// TwinCAT 3 PLC project TC3_Tester_Palet
// ProgramVersion: 3.1.4026.26
// libraries:
//   Tc2_Standard, * (Beckhoff Automation GmbH)
//   Tc2_System, * (Beckhoff Automation GmbH)
// project tree:
//   DUTs/DUTs/ E_StackAlarm.TcDUT, ST_StackCfg.TcDUT, ST_StackMem.TcDUT, ST_StackPersist.TcDUT, ST_St04Cfg.TcDUT, ST_St04_In.TcDUT, ST_St04_Out.TcDUT, ST_St05Cfg.TcDUT, ST_St05_In.TcDUT, ST_St05_Out.TcDUT, E_CylAlarm.TcDUT, E_CylFeedback.TcDUT, E_CylState.TcDUT, E_CylValve.TcDUT, ST_CylCfg.TcDUT, ST_CylMem.TcDUT, ST_CylPersist.TcDUT, E_MachineMode.TcDUT, E_NodeAlarm.TcDUT, E_NodeState.TcDUT, E_WaitCause.TcDUT, ST_ConvCfg.TcDUT, ST_ConvMem.TcDUT, ST_ConvPersist.TcDUT, E_NordSK550P_State.TcDUT, ST_NordSK550P_In.TcDUT, ST_NordSK550P_Out.TcDUT
//   POUs/POUs/FB/ FB_StackLift.TcPOU, FB_Station03_Destack.TcPOU, FB_Station11_Stack.TcPOU, FB_Station04_Press.TcPOU, FB_Station05_Tear.TcPOU, FB_CylPosMonitor.TcPOU, FB_CamAxis.TcPOU, FB_CsvLogger.TcPOU, FB_Cylinder.TcPOU, FB_RollerConveyor.TcPOU, FB_TransportNodeBase.TcPOU, FB_StationPickup.TcPOU, FB_NordSK550PP.TcPOU, TestFb.TcPOU
//   GVLs/ GVL_PERSIST.TcGVL, GVL.TcGVL, GVL_IO.TcGVL, GVL_SAFETY.TcGVL
//   / PlcTask.TcTTO
//   POUs/ PRG_Machine.TcPOU, MAIN.TcPOU

CONFIGURATION TC3_Tester_Palet
    RESOURCE PLC ON TwinCAT3
        TASK PlcTask(INTERVAL := T#10ms, PRIORITY := 20);
        PROGRAM MAIN WITH PlcTask : MAIN;
    END_RESOURCE
END_CONFIGURATION

// ---- DUTs/DUTs/E_StackAlarm.TcDUT
TYPE E_StackAlarm :
(
	ALM_STK_NONE			:= 0,

	// Wozek nie dojechal do pozycji w zadanym czasie
	ALM_STK_MOVE_TIMEOUT	:= 1,

	// Szczeki nie potwierdzily ruchu
	ALM_STK_JAW_TIMEOUT		:= 2,

	// Pozycje wpisane przez operatora nie tworza rosnacego
	// ani malejacego ciagu - dol / srodek / gora musza lezec
	// po kolei, inaczej wozek pojechalby w zla strone
	ALM_STK_POS_INVALID		:= 3,

	// Blad falownika wozka
	ALM_STK_DRIVE_FAULT		:= 4,

	// Brak wywolania M_Config
	ALM_STK_NOT_CONFIGURED	:= 5,

	// Wozek zjechal z potwierdzonej pozycji bez komendy
	ALM_STK_POSITION_LOST	:= 6
);
END_TYPE

// ---- DUTs/DUTs/ST_StackCfg.TcDUT
TYPE ST_StackCfg :
STRUCT
	// =========================================================
	// DESZTAPLARKA / SZTAPLARKA - NASTAWY NIEULOTNE
	// =========================================================
	//
	// Obie maszyny maja te sama kinematyke: wozek ze szczekami
	// jezdzacy w pionie na falowniku, z enkoderem absolutnym,
	// i trzy pozycje robocze. Rozni je tylko kolejnosc krokow.
	//
	// ---------------------------------------------------------
	// TRZY POZYCJE
	// ---------------------------------------------------------
	// Liczac od dolu, przy stosie stojacym na transporterze:
	//
	//   diPosBottom  wysokosc desek PIERWSZEJ palety od dolu
	//   diPosMiddle  wysokosc desek DRUGIEJ palety od dolu
	//   diPosTop     pozycja stosu uniesionego
	//
	// Desztaplarka chwyta na diPosMiddle - czyli pod druga
	// palete - i jedzie na diPosTop, przez co najnizsza paleta
	// zostaje na transporterze. Odklada stos na diPosBottom.
	//
	// Sztaplarka odklada trzymany stos na diPosMiddle, czyli
	// wprost na palete, ktora wlasnie przyjechala, a chwyta
	// caly stos od spodu na diPosBottom.
	//
	// Wartosci wpisuje operator z palca. Automat bazujacy
	// dopiszemy pozniej - dlatego jest kontrola poprawnosci:
	// trzy pozycje musza tworzyc ciag rosnacy albo malejacy.

	sName				: STRING(31);

	// Wartosci dobrane na maszynie. Enkoder jednoobrotowy
	// 0..65535, zero na pozycji DOLNEJ. Obie maszyny maja na
	// razie te same punkty.
	//
	// UWAGA: to sa wartosci NIEULOTNE. Wpis z deklaracji
	// obowiazuje tylko przy pierwszym pobraniu projektu albo
	// po skasowaniu danych nieulotnych. Pozniejsza zmiana tej
	// liczby w kodzie nie ruszy nastawy na sterowniku - trzeba
	// ja poprawic online albo zrobic "Reset origin".
	diPosBottom			: DINT := 0;
	diPosMiddle			: DINT := 16000;
	diPosTop			: DINT := 24000;

	// Okno, w ktorym uznajemy pozycje za osiagnieta
	diWindow			: DINT := 20;

	// Odleglosc, od ktorej zwalniamy do predkosci dojazdowej
	diSlowZone			: DINT := 300;

	// TRUE = rosnaca wartosc enkodera odpowiada jezdzie
	// napedem DO PRZODU
	xIncreaseIsForward	: BOOL := TRUE;


	// ---------------------------------------------------------
	// PREDKOSCI I CZASY
	// ---------------------------------------------------------

	lrFreqFast			: LREAL := 35.0;
	lrFreqSlow			: LREAL := 10.0;
	lrFreqManual		: LREAL := 8.0;

	// Czas, w ktorym wozek musi dojechac do pozycji
	tMoveWatchdog		: TIME := T#15S;

	// Uspokojenie po dojezdzie, zanim ruszymy szczekami
	tSettle				: TIME := T#200MS;


	// ---------------------------------------------------------
	// STOS
	// ---------------------------------------------------------
	//
	// Na razie stala liczba palet w stosie. Czujnik wykrywajacy,
	// ze wszystkie palety zostaly wydane, dojdzie pozniej -
	// wtedy ta wartosc bedzie tylko wartoscia oczekiwana.

	nStackSize			: INT := 15;

END_STRUCT
END_TYPE

// ---- DUTs/DUTs/ST_StackMem.TcDUT
TYPE ST_StackMem :
STRUCT
	// =========================================================
	// PAMIEC DESZTAPLARKI / SZTAPLARKI - ZMIENNE NIEULOTNE
	// =========================================================
	//
	// Po zaniku zasilania maszyna musi wiedziec, ile palet
	// zostalo w stosie i ile wisi na szczekach. Bez tego
	// operator musialby rozladowac stacje recznie.

	// Stos dojechal na stacje i zostal potwierdzony czujnikami
	xStackArrived	: BOOL;

	// DESZTAPLARKA: ile palet zostalo do wydania, wliczajac te,
	// ktora aktualnie lezy na transporterze
	nRemaining		: INT;

	// SZTAPLARKA: ile palet wisi na szczekach
	nHeld			: INT;

	// Szczeki trzymaja ladunek - po zaniku zasilania nie wolno
	// ich otworzyc bez sprowadzenia wozka na pozycje odkladania
	xJawsLoaded		: BOOL;

	// Ostatnia znana pozycja enkodera, zapisywana na biezaco.
	// Po starcie porownujemy ja z odczytem: jesli sie zgadza,
	// enkoder utrzymal wartosc przez zanik zasilania i NIE ma
	// potrzeby bazowania. Jesli nie - kod sam to zglosi.
	diLastPos		: DINT;

	// TRUE = po starcie odczyt enkodera nie zgodzil sie
	// z zapamietanym. Trzeba zbazowac pozycje dolna.
	xNeedHoming		: BOOL;

END_STRUCT
END_TYPE

// ---- DUTs/DUTs/ST_StackPersist.TcDUT
TYPE ST_StackPersist :
STRUCT
	Cfg		: ST_StackCfg;
	Mem		: ST_StackMem;
END_STRUCT
END_TYPE

// ---- DUTs/DUTs/ST_St04Cfg.TcDUT
TYPE ST_St04Cfg :
STRUCT
	// =========================================================
	// STACJA 4 - TEST SCISKANIA, NASTAWY NIEULOTNE
	// =========================================================
	//
	// Test toczy sie na JADACEJ palecie. Rolki dociskowe kreca
	// sie caly czas, a silowniki napieraja na deski w trakcie
	// przejazdu. Dlatego przerwanie uniewaznia wynik -
	// aConv[4].Cfg.xNokOnInterrupt musi byc TRUE.

	// ---------------------------------------------------------
	// CZUJNIK WSTEPNY
	// ---------------------------------------------------------
	//
	// Czujnik przed stacja, od ktorego liczy sie czas do wysuwu
	// silownikow. Na dzien pisania kodu jeszcze nie zamontowany.
	//
	// xPreSensorInstalled = FALSE: czasowka startuje od chwili
	// ruszenia palety z poprzedniej stacji (tEntryToUpper).
	// Po montazu wystarczy przelaczyc bit - kod sie nie zmienia.

	xPreSensorInstalled	: BOOL := FALSE;

	// TRUE = logika odwrocona, tak jak czujniki koncowe
	// (0 na wejsciu = czujnik cos widzi)
	xPreSensorInverted	: BOOL := TRUE;


	// ---------------------------------------------------------
	// CZASY SEKWENCJI
	// ---------------------------------------------------------

	// Od czujnika wstepnego do wysuwu silownikow GORNYCH
	tPreToUpper			: TIME := T#500MS;

	// To samo, gdy czujnika wstepnego jeszcze nie ma -
	// liczone od rozpoczecia wjazdu
	tEntryToUpper		: TIME := T#3S;

	// Od wysuwu gornych do wysuwu DOLNYCH.
	// Gorne ida pierwsze, zeby dolne nie uniosly palety,
	// ale odstep ma byc symboliczny - dociski maja isc razem.
	tUpperToLower		: TIME := T#100MS;

	// Watchdog calej operacji
	tOpWatchdog			: TIME := T#60S;


	// ---------------------------------------------------------
	// ROLKI DOCISKOWE
	// ---------------------------------------------------------
	//
	// Falownik 3. Rolki na koncach silownikow gornych sa
	// napedzane, zeby paleta nie utknela pod dociskiem.

	lrRollerFreq		: LREAL := 25.0;

END_STRUCT
END_TYPE

// ---- DUTs/DUTs/ST_St04_In.TcDUT
TYPE ST_St04_In :
STRUCT
	// =========================================================
	// STACJA 4 - SYGNALY WEJSCIOWE
	// =========================================================

	// Czujnik wstepny - jeszcze niepodlinkowany.
	// Do czasu montazu zostawic Cfg.xPreSensorInstalled = FALSE.
	xPreSensRaw		: BOOL := TRUE;

	// Przetworniki polozenia IO-Link, po jednym na KAZDY
	// silownik, mimo ze zawory steruja grupami:
	//   1..3  dolne
	//   4..6  gorne od szerokich desek
	//   7..8  gorne od waskich desek
	adiCylPos		: ARRAY[1..8] OF DINT;

END_STRUCT
END_TYPE

// ---- DUTs/DUTs/ST_St04_Out.TcDUT
TYPE ST_St04_Out :
STRUCT
	// =========================================================
	// STACJA 4 - CEWKI ZAWOROW
	// =========================================================
	//
	// Mapowanie w MAIN wg opisu wyjsc:
	//   xLowerExtend        -> GVL.OUTPUTS[4]   dolne wysun
	//   xLowerRetract       -> GVL.OUTPUTS[3]   dolne cofnij
	//   xUpperWideExtend    -> GVL.OUTPUTS[7]   gorne zewnetrzne
	//                                           i srodkowa wysun
	//   xUpperWideRetract   -> GVL.OUTPUTS[2]   te same cofnij
	//   xUpperNarrowExtend  -> GVL.OUTPUTS[5]   gorne srodkowe wysun
	//   xUpperNarrowRetract -> GVL.OUTPUTS[6]   gorne srodkowe cofnij
	//
	// [?] Opis wyjsc 2/7 i 5/6 nazywa obie grupy "srodkowymi".
	// Przyjete: 7/2 to trzy silowniki od szerokich desek,
	// 5/6 to dwa od waskich. Do potwierdzenia na maszynie -
	// zamiana dotyczy wylacznie mapowania w MAIN, nie kodu stacji.

	xLowerExtend		: BOOL;
	xLowerRetract		: BOOL;

	xUpperWideExtend	: BOOL;
	xUpperWideRetract	: BOOL;

	xUpperNarrowExtend	: BOOL;
	xUpperNarrowRetract	: BOOL;

END_STRUCT
END_TYPE

// ---- DUTs/DUTs/ST_St05Cfg.TcDUT
TYPE ST_St05Cfg :
STRUCT
	// =========================================================
	// STACJA 5 - TEST ROZRYWANIA, NASTAWY NIEULOTNE
	// =========================================================
	//
	// Czasy samych ruchow silownikow siedza w ich wlasnych
	// rekordach (GVL_PERSIST.aCyl). Tutaj sa tylko czasy
	// nalezace do SEKWENCJI stacji.

	// Od potwierdzenia palety na blokadzie do podniesienia szczek
	tDetectToLift		: TIME := T#500MS;

	// Od zamkniecia szczek do rozpoczecia rozrywania
	tJawsToPull			: TIME := T#300MS;

	// Watchdog calej operacji testu
	tOpWatchdog			: TIME := T#60S;

	// UWAGA: blokada NIE podnosi sie na czasowke. Idzie w gore
	// w chwili, gdy z poprzedniej stacji rusza paleta - wtedy
	// nikt jej nie stoi na drodze, a czasu na podniesienie jest
	// tyle, ile trwa przejazd. Czas ruchu samej blokady i jego
	// watchdog siedza w GVL_PERSIST.aCyl.

END_STRUCT
END_TYPE

// ---- DUTs/DUTs/ST_St05_In.TcDUT
TYPE ST_St05_In :
STRUCT
	// =========================================================
	// STACJA 5 - SYGNALY WEJSCIOWE
	// =========================================================
	//
	// Cale mapowanie z GVL siedzi w jednym miejscu w MAIN.
	// Blok stacji nie siega do GVL bezposrednio.

	// Blokada punktu zatrzymania - czujniki gorny i dolny
	xBlockUpSw		: BOOL;
	xBlockDownSw	: BOOL;

	// Silownik podnoszenia szczek - czujniki po obu stronach
	xJawLiftUpSw	: BOOL;
	xJawLiftDownSw	: BOOL;

	// Czujniki otwarcia szczek. Trzy pary po dwa silowniki,
	// para obsluguje jedna dolna deske palety. Para jest
	// otwarta dopiero gdy OBA silowniki zglaszaja otwarcie -
	// tylko wtedy wolno wjechac i wyjechac paleta.
	axJawOpenSw		: ARRAY[1..3, 1..2] OF BOOL;

	// Przetworniki polozenia silownikow rozrywajacych,
	// indeksowane NUMEREM SILOWNIKA 1..6 (nie numerem zaworu)
	adiPullPos		: ARRAY[1..6] OF DINT;

END_STRUCT
END_TYPE

// ---- DUTs/DUTs/ST_St05_Out.TcDUT
TYPE ST_St05_Out :
STRUCT
	// =========================================================
	// STACJA 5 - CEWKI ZAWOROW
	// =========================================================
	//
	// Mapowanie w MAIN:
	//   xBlockExtend    -> FestoValves_1[6,1]   blokada w gore
	//   xBlockRetract   -> FestoValves_1[6,2]   blokada w dol
	//   xJawLiftExtend  -> FestoValves_1[7,1]   szczeki w gore
	//   xJawLiftRetract -> FestoValves_1[7,2]   szczeki w dol
	//   axJawClose[1]   -> FestoValves_1[1,1]   szczeki lewe
	//   axJawClose[2]   -> FestoValves_1[2,1]   szczeki srodkowe
	//   axJawClose[3]   -> FestoValves_1[3,1]   szczeki prawe
	//
	// Silowniki rozrywajace - UWAGA, numer zaworu nie jest
	// numerem silownika:
	//   silownik 1 -> FestoValves_2[4,2] gora / [4,1] dol
	//   silownik 2 -> FestoValves_2[3,2] gora / [3,1] dol
	//   silownik 3 -> FestoValves_2[1,2] gora / [1,1] dol
	//   silownik 4 -> FestoValves_2[2,2] gora / [2,1] dol
	//   silownik 5 -> FestoValves_2[5,2] gora / [5,1] dol
	//   silownik 6 -> FestoValves_2[6,2] gora / [6,1] dol
	//
	// Tablice ponizej sa indeksowane NUMEREM SILOWNIKA.

	xBlockExtend	: BOOL;
	xBlockRetract	: BOOL;

	xJawLiftExtend	: BOOL;
	xJawLiftRetract	: BOOL;

	// TRUE = szczeki zamkniete (zawor monostabilny)
	axJawClose		: ARRAY[1..3] OF BOOL;

	axPullUp		: ARRAY[1..6] OF BOOL;
	axPullDown		: ARRAY[1..6] OF BOOL;

END_STRUCT
END_TYPE

// ---- DUTs/DUTs/E_CylAlarm.TcDUT
TYPE E_CylAlarm :
(
	ALM_CYL_NONE				:= 0,

	// Nie potwierdzil wysuwu w czasie tExtendWatchdog
	ALM_CYL_EXTEND_TIMEOUT		:= 1,

	// Nie potwierdzil wsuwu w czasie tRetractWatchdog
	ALM_CYL_RETRACT_TIMEOUT		:= 2,

	// Obie krancowki aktywne jednoczesnie
	ALM_CYL_BOTH_SWITCHES		:= 3,

	// Przetwornik nie zostal zbazowany, a progi sa uzywane
	ALM_CYL_NOT_ZEROED			:= 4,

	// Zejscie z potwierdzonego polozenia bez komendy
	ALM_CYL_POSITION_LOST		:= 5,

	// Brak wywolania M_Config
	ALM_CYL_NOT_CONFIGURED		:= 6
);
END_TYPE

// ---- DUTs/DUTs/E_CylFeedback.TcDUT
TYPE E_CylFeedback :
(
	// Brak sprzezenia - ruch wylacznie na czasowkach
	CYLFB_NONE		:= 0,

	// Krancowki na jednym albo obu koncach
	CYLFB_SWITCHES	:= 1,

	// Przetwornik polozenia IO-Link, wartosc bezwzgledna DINT.
	// Polozenia koncowe to progi nastawiane przez operatora,
	// a nie zdarzenia dwustanowe.
	CYLFB_ANALOG	:= 2,

	// Sprzezenie podawane z zewnatrz przez stacje.
	// Uzywane tam, gdzie jeden zawor steruje GRUPA silownikow,
	// a pomiar jest indywidualny - stacja 4. Stacja agreguje
	// wskazania FB_CylPosMonitor i podaje wynik na wejscia
	// xFbExtIn / xFbRetIn.
	CYLFB_EXTERNAL	:= 3
);
END_TYPE

// ---- DUTs/DUTs/E_CylState.TcDUT
TYPE E_CylState :
(
	// Polozenie nieznane - po starcie, przed pierwsza komenda
	// albo po powrocie z trybu recznego
	CYL_UNKNOWN		:= 0,

	CYL_RETRACTED	:= 10,
	CYL_EXTENDING	:= 20,
	CYL_EXTENDED	:= 30,
	CYL_RETRACTING	:= 40,

	CYL_MANUAL		:= 70,
	CYL_ALARM		:= 90
);
END_TYPE

// ---- DUTs/DUTs/E_CylValve.TcDUT
TYPE E_CylValve :
(
	// Zawor monostabilny, jedna cewka.
	// TRUE = wysuniety, FALSE = wycofany sprezyna.
	// Przyklad: szczeki stacji 5, FestoValves_1[1..3, 1]
	CYLV_SINGLE			:= 0,

	// Zawor bistabilny, dwie cewki wykluczajace sie
	CYLV_DOUBLE			:= 1,

	// Zawor 3-polozeniowy. Wysuw i cofniecie po wlasnej cewce,
	// oba wyjscia zdjete = polozenie spoczynkowe (srodkowe).
	CYLV_3POS_MID		:= 2,

	// Zawor 3-polozeniowy, w ktorym cofniecie realizuje
	// zdjecie OBU cewek
	CYLV_3POS_OFF_RET	:= 3
);
END_TYPE

// ---- DUTs/DUTs/ST_CylCfg.TcDUT
TYPE ST_CylCfg :
STRUCT
	// =========================================================
	// NASTAWY SILOWNIKA - ZMIENNE NIEULOTNE
	// =========================================================
	//
	// Edytowalne przez operatora z HMI. Kod ich nie zapisuje -
	// jedyny wyjatek to bazowanie przetwornika, ktore siedzi
	// w ST_CylMem.

	sName				: STRING(31);

	eValve				: E_CylValve;
	eFeedback			: E_CylFeedback;


	// ---------------------------------------------------------
	// CZASOWKI
	// ---------------------------------------------------------

	// Opoznienie wysterowania zaworu po otrzymaniu komendy.
	// Sluzy do rozjezdzania w czasie silownikow, ktore nie
	// moga ruszyc razem - np. gorne przed dolnymi na stacji 4.
	tExtendDelay		: TIME := T#0MS;
	tRetractDelay		: TIME := T#0MS;

	// Czas, w ktorym ruch musi sie zakonczyc
	tExtendWatchdog		: TIME := T#3S;
	tRetractWatchdog	: TIME := T#3S;

	// Watchdog wylaczalny osobno dla kazdego kierunku.
	// Silownik bez krancowki na jednym koncu nie ma jak
	// potwierdzic dojazdu - wtedy watchdog w tym kierunku
	// musi byc wylaczony.
	xExtendWdEnabled	: BOOL := TRUE;
	xRetractWdEnabled	: BOOL := TRUE;


	// ---------------------------------------------------------
	// SPRZEZENIE OD POLOZENIA
	// ---------------------------------------------------------
	//
	// Obserwacje polozenia koncowego mozna wylaczyc OSOBNO dla
	// kazdego kierunku i zastapic czasowka. To jest tryb pracy
	// z uszkodzonym czujnikiem: PLC uznaje ruch za wykonany po
	// uplywie czasu.

	xExtendFbEnabled	: BOOL := TRUE;
	xRetractFbEnabled	: BOOL := TRUE;

	tExtendSubst		: TIME := T#1S;
	tRetractSubst		: TIME := T#1S;

	// Czas stabilnego stanu potrzebny do uznania niezgodnosci
	// krancowek za rzeczywista
	tSettle				: TIME := T#500MS;


	// ---------------------------------------------------------
	// PROGI PRZETWORNIKA IO-LINK (tylko CYLFB_ANALOG)
	// ---------------------------------------------------------
	//
	// Wszystkie progi liczone WZGLEDEM punktu bazowania.
	// Znak dodatni zawsze w kierunku wysuwu - jesli przetwornik
	// liczy odwrotnie, ustawic xInvertPos.
	//
	// Stacja 4 bazuje na silowniku WYSUNIETYM z paleta,
	// stacja 5 na silowniku WYCOFANYM. Dlatego progi moga
	// byc ujemne i nie jest to blad.

	xInvertPos			: BOOL := FALSE;

	// Ponizej tej wartosci uznajemy silownik za wycofany
	diPosRetracted		: DINT := 100;

	// Powyzej tej wartosci uznajemy silownik za wysuniety
	diPosExtended		: DINT := 1000;

	// Przekroczenie = deska pekla albo odpadla.
	// To jest WYNIK TESTU, nie alarm silownika.
	diPosLimit			: DINT := 2000;

	// Powyzej tej wartosci zaczynamy liczyc czas trzymania
	// nacisku (stacja 5)
	diPosHoldStart		: DINT := 1500;
	tHold				: TIME := T#2S;

END_STRUCT
END_TYPE

// ---- DUTs/DUTs/ST_CylMem.TcDUT
TYPE ST_CylMem :
STRUCT
	// =========================================================
	// PAMIEC SILOWNIKA - ZMIENNE NIEULOTNE
	// =========================================================

	// Wskazanie surowe przetwornika w punkcie bazowania.
	// Zapisuje je procedura M_Zero w trybie recznym.
	diZeroOffset	: DINT;

	// FALSE = przetwornik nigdy nie byl bazowany, progi
	// polozenia nic nie znacza
	xZeroed			: BOOL;

END_STRUCT
END_TYPE

// ---- DUTs/DUTs/ST_CylPersist.TcDUT
TYPE ST_CylPersist :
STRUCT
	Cfg		: ST_CylCfg;
	Mem		: ST_CylMem;
END_STRUCT
END_TYPE

// ---- DUTs/DUTs/E_MachineMode.TcDUT
TYPE E_MachineMode :
(
	// Maszyna zatrzymana - zadna sekwencja nie pracuje
	MODE_STOP		:= 0,

	// Praca automatyczna
	MODE_AUTO		:= 1,

	// Praca reczna - sterowanie pojedynczymi elementami,
	// dozwolony ruch w obu kierunkach
	MODE_MANUAL		:= 2,

	// Praca krokowa - sekwencja czeka na potwierdzenie
	// operatora przed kazdym krokiem
	MODE_STEP		:= 3,

	// Bazowanie / odstawianie do pozycji startowej
	MODE_HOME		:= 4
);
END_TYPE

// ---- DUTs/DUTs/E_NodeAlarm.TcDUT
TYPE E_NodeAlarm :
(
	ALM_NONE					:= 0,

	// Ladunek nie dojechal w czasie tInfeedWatchdog
	ALM_INFEED_TIMEOUT			:= 1,

	// Ladunek nie zjechal w czasie tOutfeedWatchdog
	ALM_OUTFEED_TIMEOUT			:= 2,

	// Pamiec mowi "pusto", czujniki widza ladunek
	ALM_UNEXPECTED_LOAD			:= 3,

	// Pamiec mowi "zajete", czujniki nie widza nic
	ALM_LOAD_LOST				:= 4,

	// Czujniki nie zgadzaja sie ze soba po zatrzymaniu
	ALM_SENSOR_DISAGREE			:= 5,

	// Blad falownika
	ALM_DRIVE_FAULT				:= 6,

	// Falownik nie potwierdzil ruchu mimo zadania
	ALM_DRIVE_NO_FEEDBACK		:= 7,

	// Wyczerpano liczbe prob wznowienia przerwanego przejazdu
	ALM_RESUME_FAILED			:= 8,

	// Brak wywolania M_Config - wezel nie ma parametrow
	ALM_NOT_CONFIGURED			:= 9,

	// Operacja technologiczna stacji zglosila blad
	ALM_OPERATION_FAILED		:= 10
);
END_TYPE

// ---- DUTs/DUTs/E_NodeState.TcDUT
TYPE E_NodeState :
(
	// Stan poczatkowy - weryfikacja pamieci wzgledem czujnikow
	NODE_INIT		:= 0,

	// Wezel pusty, gotowy przyjac ladunek
	NODE_EMPTY		:= 10,

	// Ladunek wjezdza na wezel
	NODE_INFEED		:= 20,

	// Wykryto pozycje koncowa, trwa czasowka do zatrzymania
	NODE_STOP_DELAY	:= 30,

	// Ladunek stoi, brak operacji technologicznej
	NODE_OCCUPIED	:= 40,

	// Trwa operacja technologiczna stacji
	NODE_BUSY		:= 50,

	// Wydawanie ladunku na nastepny wezel
	NODE_OUTFEED	:= 60,

	// Praca reczna
	NODE_MANUAL		:= 70,

	// Pamiec nie zgadza sie z czujnikami - wymagana decyzja operatora
	NODE_VERIFY		:= 80,

	// Alarm - ruch zablokowany do czasu resetu
	NODE_ALARM		:= 90
);
END_TYPE

// ---- DUTs/DUTs/E_WaitCause.TcDUT
TYPE E_WaitCause :
(
	// =========================================================
	// JEDNOZNACZNA PRZYCZYNA POSTOJU
	// =========================================================
	//
	// W kazdym cyklu wezel ustawia DOKLADNIE JEDNA przyczyne.
	// Jesli wezel stoi, ta zmienna mowi czego brakuje - bez
	// koniecznosci wchodzenia w kod.

	WAIT_NONE				:= 0,

	// --- warunki wlasne wezla ---
	WAIT_NO_SAFETY			:= 1,	// STO / lancuch bezpieczenstwa
	WAIT_NOT_AUTO			:= 2,	// tryb inny niz AUTO
	WAIT_ALARM_ACTIVE		:= 3,	// alarm wlasny
	WAIT_STATE_UNVERIFIED	:= 4,	// pamiec wymaga potwierdzenia
	WAIT_NO_LOAD			:= 5,	// pusto, nie ma czego wydac
	WAIT_OPERATION_BUSY		:= 6,	// trwa operacja technologiczna
	WAIT_DRIVE_NOT_READY	:= 7,	// falownik niegotowy
	WAIT_DRIVE_FAULT		:= 8,	// blad falownika
	WAIT_STEP_ACK			:= 9,	// tryb krokowy - brak potwierdzenia
	WAIT_NOT_CONFIGURED		:= 10,	// brak M_Config
	WAIT_STATION_NOT_READY	:= 11,	// mechanika stacji nie w pozycji
	WAIT_TRANSFER_HOLD		:= 12,	// zdjete reczne zezwolenie na przejazd
	WAIT_PICKUP				:= 13,	// czeka na odbior przez operatora

	// --- warunki nastepnego wezla ---
	WAIT_NEXT_NOT_LINKED	:= 20,	// nie podpieto nastepnika
	WAIT_NEXT_OCCUPIED		:= 21,	// nastepnik zajety
	WAIT_NEXT_ALARM			:= 22,	// nastepnik w alarmie
	WAIT_NEXT_UNVERIFIED	:= 23,	// nastepnik wymaga weryfikacji
	WAIT_NEXT_NOT_AUTO		:= 24,	// nastepnik nie w AUTO
	WAIT_NEXT_NO_SAFETY		:= 25,	// nastepnik bez zezwolenia
	WAIT_NEXT_BUSY			:= 26,	// nastepnik w trakcie operacji

	// --- warunki poprzedniego wezla ---
	WAIT_PREV_NOT_READY		:= 30
);
END_TYPE

// ---- DUTs/DUTs/ST_ConvCfg.TcDUT
TYPE ST_ConvCfg :
STRUCT
	// =========================================================
	// NASTAWY TRANSPORTERA - ZMIENNE NIEULOTNE
	// =========================================================
	//
	// Caly ten rekord jest edytowalny przez operatora z HMI.
	// Instancja lezy w GVL_PERSIST.aConv[n], FB dostaje na nia
	// wskaznik przez M_Config. Nic w tej strukturze nie jest
	// modyfikowane przez kod - tylko przez operatora.

	// Opis wezla na HMI
	sName				: STRING(31);


	// ---------------------------------------------------------
	// NAPED
	// ---------------------------------------------------------

	// Czestotliwosc w pracy automatycznej [Hz]
	lrFreqAuto			: LREAL := 30.0;

	// Czestotliwosc w pracy recznej [Hz]
	lrFreqManual		: LREAL := 15.0;

	// Trwale odwrocenie kierunku obrotow.
	// Dla silnikow podlaczonych odwrotnie - zamiast przekladac
	// fazy, odwracamy bit w jednym miejscu.
	xInvertDirection	: BOOL := FALSE;

	// Opoznienie zatrzymania po wykryciu pozycji przez czujniki
	tStopDelay			: TIME := T#150MS;


	// ---------------------------------------------------------
	// CZUJNIKI
	// ---------------------------------------------------------
	//
	// Czujniki pracuja w logice odwroconej: sygnal 1 = wolne,
	// sygnal 0 = cos widac. Obecnosc w pozycji koncowej to
	// zero z OBU czujnikow.
	//
	// Wylaczenie czujnika = serwis uznal go za uszkodzony,
	// jego sygnal jest ignorowany. Wylaczenie OBU przelacza
	// wezel w tryb czasowkowy (patrz tBlindTravel).

	xSensor1Enabled		: BOOL := TRUE;
	xSensor2Enabled		: BOOL := TRUE;

	// Polaryzacja czujnikow.
	// TRUE  - logika odwrocona: 0 = czujnik cos widzi (maszyna docelowa)
	// FALSE - logika wprost:    1 = czujnik cos widzi (wersja testowa)
	xSensorsInverted	: BOOL := TRUE;

	// Czas stabilnego stanu, po ktorym uznajemy niezgodnosc
	// czujnikow albo niezgodnosc pamieci za rzeczywista
	tSensorSettle		: TIME := T#1S;


	// ---------------------------------------------------------
	// CZASY PRZEJAZDU
	// ---------------------------------------------------------

	// Watchdog wjazdu - po tym czasie ladunek MUSI byc
	// w pozycji koncowej, inaczej alarm
	tInfeedWatchdog		: TIME := T#20S;

	// Watchdog wyjazdu - po tym czasie ladunek MUSI zejsc
	// z pola czujnikow, inaczej alarm
	tOutfeedWatchdog	: TIME := T#20S;

	// Czas przejazdu w trybie bez czujnikow. Liczony od
	// jednoczesnego ruszenia obu transporterow.
	tBlindTravel		: TIME := T#6S;

	// Czas potwierdzenia, ze ladunek naprawde zjechal
	tClearDelay			: TIME := T#500MS;


	// ---------------------------------------------------------
	// ZACHOWANIE
	// ---------------------------------------------------------

	// Operacja technologiczna stacji wlaczona.
	// FALSE = stacja realizuje wylacznie przejazd.
	xStationEnabled		: BOOL := TRUE;

	// Zgoda na przejazd bez zatrzymania, gdy na wezle nie ma
	// nic do zrobienia a nastepnik jest gotowy
	xAllowPassThrough	: BOOL := TRUE;

	// Przerwanie operacji unieważnia wynik testu.
	//
	// TRUE  - grzyb, kurtyna, przeciazenie napedu, zanik
	//         zasilania w trakcie testu oznaczaja, ze wyniku
	//         nie da sie juz uznac za wiarygodny: paleta idzie
	//         na odrzut i nie jest badana ponownie.
	//         Ustawic na stacjach 4 i 6.
	//
	// FALSE - po ustapieniu przyczyny mozna kontynuowac albo
	//         powtorzyc cykl od poczatku. Pozostale stacje.
	xNokOnInterrupt		: BOOL := FALSE;

	// Ile razy maszyna sprobuje sama dokonczyc przerwany
	// przejazd po resecie operatora
	nResumeRetries		: INT := 1;

	// Odbior przez operatora potwierdzany przyciskiem.
	// FALSE = miejsce uznajemy za wolne po tPickupTimeout
	// od zniknieca ladunku z czujnikow (stacje 13 i 16).
	xPickupByButton		: BOOL := TRUE;
	tPickupTimeout		: TIME := T#10S;

END_STRUCT
END_TYPE

// ---- DUTs/DUTs/ST_ConvMem.TcDUT
TYPE ST_ConvMem :
STRUCT
	// =========================================================
	// PAMIEC STANU TRANSPORTERA - ZMIENNE NIEULOTNE
	// =========================================================
	//
	// To NIE sa nastawy. Ta struktura przezywa zanik zasilania
	// i po starcie maszyna wie, gdzie stoja palety.
	//
	// UWAGA: kazda zmiana pola w tej strukturze musi ustawic
	// xPersistDirty w wezle, zeby menedzer zapisal dane na
	// dysk. Bez tego przy zaniku zasilania stracimy obraz.

	// Obraz obecnosci ladunku. Ustawiany na TRUE w chwili
	// ROZPOCZECIA wjazdu, kasowany dopiero po potwierdzonym
	// zjezdzie - w trakcie przejazdu oba wezly sa "zajete",
	// bo paleta fizycznie lezy na obu.
	xLoadPresent		: BOOL;

	// FALSE = pamiec rozjechala sie z czujnikami i operator
	// musi rozstrzygnac stan. Wezel nie ruszy do tego czasu.
	xStateVerified		: BOOL := TRUE;

	// Przejazd zostal przerwany (STO, zanik zasilania,
	// watchdog, zaciecie). Po resecie maszyna sprobuje
	// dokonczyc ruch od tej fazy.
	xTransferAborted	: BOOL;
	eAbortedPhase		: E_NodeState;

	// Licznik prob automatycznego wznowienia
	nResumeCount		: INT;

	// Operacja technologiczna dla lezacego ladunku zostala
	// dokonczona. Bez tego po restarcie w polowie testu paleta
	// wyjechalaby nieprzebadana i zaliczona jako dobra.
	xOperationDone		: BOOL;

	// Operacja zostala przerwana w polowie - grzyb, kurtyna,
	// przeciazenie napedu, zanik zasilania. Na stacjach
	// z Cfg.xNokOnInterrupt oznacza to odrzut palety.
	xOperationInterrupted	: BOOL;

	// Werdykt dla ladunku lezacego na wezle.
	// TRUE = paleta odrzucona, nie realizujemy dla niej
	// zadnych dalszych testow ani etykietowania.
	xLoadNok			: BOOL;

	// Numer sztuki - do sledzenia palety przez maszyne
	nLoadId				: UDINT;

END_STRUCT
END_TYPE

// ---- DUTs/DUTs/ST_ConvPersist.TcDUT
TYPE ST_ConvPersist :
STRUCT
	// Nastawy operatora
	Cfg		: ST_ConvCfg;

	// Pamiec stanu maszyny
	Mem		: ST_ConvMem;
END_STRUCT
END_TYPE

// ---- DUTs/DUTs/E_NordSK550P_State.TcDUT
TYPE E_NordSK550P_State :
(
    NORD_STATE_NOT_READY,
    NORD_STATE_SWITCH_ON_DISABLED,
    NORD_STATE_READY_TO_SWITCH_ON,
    NORD_STATE_SWITCHED_ON,
    NORD_STATE_OPERATION_ENABLED,
    NORD_STATE_QUICK_STOP_ACTIVE,
    NORD_STATE_FAULT_REACTION_ACTIVE,
    NORD_STATE_FAULT,
    NORD_STATE_UNKNOWN
);
END_TYPE

// ---- DUTs/DUTs/ST_NordSK550P_In.TcDUT
TYPE ST_NordSK550P_In :
STRUCT
    // 0x6061
    byModeDisplay : USINT;

    // 0x6041
    wStatusWord : UINT;

    // 0x6043
    iVelocityDemand : INT;
END_STRUCT
END_TYPE

// ---- DUTs/DUTs/ST_NordSK550P_Out.TcDUT
TYPE ST_NordSK550P_Out :
STRUCT
    // 0x6060
    byModeOfOperation : USINT;

    // 0x6040
    wControlWord : UINT;

    // 0x60FF
    diTargetVelocity : INT;
END_STRUCT
END_TYPE

// ---- GVLs/GVL_PERSIST.TcGVL
VAR_GLOBAL PERSISTENT
	// =========================================================
	// ZMIENNE NIEULOTNE WARSTWY TRANSPORTU
	// =========================================================
	//
	// Indeks = numer stacji wg ZALOZENIA.md:
	//   1  zaladunek stosow            9  transporter lancuchowy
	//   2  bufor stosow               10  stacja przekierowujaca
	//   3  desztaplarka               11  sztaplarka
	//   4  test sciskania             12  bufor stosow (wyjscie)
	//   5  test rozrywania            13  wyjscie stosow OK
	//   6  pomiar laserowy            14  bufor odrzutu
	//   7  etykietowanie              15  bufor odrzutu
	//   8  stacja rozjazdowa          16  odbior palet NOK
	//
	// Cfg - nastawy operatora, kod ich nie zmienia.
	// Mem - obraz stanu maszyny, kod je zmienia i ustawia
	//       xPersistDirty, zeby menedzer zapisal je na dysk.
	//
	// UWAGA: wartosci poczatkowe z ST_ConvCfg sa brane pod
	// uwage TYLKO przy pierwszym pobraniu projektu. Pozniejsza
	// zmiana wartosci domyslnej w kodzie nie zmieni nastaw
	// na sterowniku - trzeba je poprawic z HMI albo wykonac
	// "Reset origin".

	aConv	: ARRAY[1..16] OF ST_ConvPersist;


	// =========================================================
	// SILOWNIKI I MONITORY POLOZENIA
	// =========================================================
	//
	// Wspolna tablica dla zaworow i dla osobnych pomiarow -
	// obie korzystaja z tego samego rekordu nastaw.
	//
	// Przydzial indeksow (do uzupelnienia przy pisaniu stacji):
	//    1.. 3  stacja 4  grupy zaworow: dolne, gorne srodkowe,
	//                     gorne zewnetrzne + srodkowa
	//    4..11  stacja 4  monitory polozenia 8 silownikow
	//   12..14  stacja 5  szczeki lewe / srodkowe / prawe
	//   15      stacja 5  blokada punktu zatrzymania
	//   16      stacja 5  podnoszenie szczek
	//   17..22  stacja 5  silowniki rozrywajace 1..6
	//   23      stacja 8  podnoszenie rolek
	//   24      stacja 10 podnoszenie rolek
	//   25..32  zapas

	aCyl	: ARRAY[1..32] OF ST_CylPersist;


	// =========================================================
	// NASTAWY SEKWENCJI STACJI
	// =========================================================

	St04	: ST_St04Cfg;
	St05	: ST_St05Cfg;


	// =========================================================
	// DESZTAPLARKA I SZTAPLARKA
	// =========================================================
	//
	// Ta sama struktura dla obu - rozni je tylko sekwencja.
	// Szczeki maja wlasne rekordy w aCyl:
	//   25  szczeki desztaplarki (stacja 3)
	//   26  szczeki sztaplarki   (stacja 11)

	St03	: ST_StackPersist;
	St11	: ST_StackPersist;

END_VAR

// ---- GVLs/GVL.TcGVL
VAR_GLOBAL
	
	NORD_DRIVE_IN AT %I* : ARRAY[1..20] OF ST_NordSK550P_In;
	NORD_DRIVE_OUT AT %Q* : ARRAY[1..20] OF ST_NordSK550P_Out;
	IO_Destaker_Act_Pos 	AT %I* : DINT;
	IO_Staker_Act_Pos 	AT %I* : DINT;
	
	FestoValves_1  AT %Q* : ARRAY[1..8, 1..2] OF BOOL;
	FestoValves_2  AT %Q* : ARRAY[1..8, 1..2] OF BOOL;
	
	
	INPUTS AT  %I* : ARRAY[1..300] OF BOOL;
	OUTPUTS AT  %Q* : ARRAY[1..300] OF BOOL;
	
	
	
END_VAR

// ---- GVLs/GVL_IO.TcGVL
VAR_GLOBAL

END_VAR

// ---- GVLs/GVL_SAFETY.TcGVL
VAR_GLOBAL
	Q_SafetyEnable AT %Q* : BOOL := TRUE;
	Q_SafetyReset AT %Q* : BOOL; 
	
	xSTO AT %I* : BOOL;
	xAir AT %I* : BOOL;
	xResetCmd AT %I* : BOOL;
	
END_VAR

// ---- POUs/MAIN.TcPOU
PROGRAM MAIN
// =============================================================
// TEST RUCHU TRANSPORTEROW
// =============================================================
//
// Proba na maszynie: jedna paleta idzie trasa, w kazdym kroku
// pracuje PARA transporterow - ten, z ktorego paleta zjezdza,
// i ten, na ktory wjezdza.
//
// -------------------------------------------------------------
// CZUJNIKI
// -------------------------------------------------------------
// Podpiete czujniki koncza przejazd zamiast czasowki.
//
//   xUseSensors   = FALSE  wracamy na same czasowki, jak dotad
//   xStepWatchdog = FALSE  krok czeka na czujnik BEZ KONCA
//
// Na czas recznego wyzwalania czujnikow watchdog jest WYLACZONY:
// zaden krok nie przeskoczy sam, dopoki nie podasz sygnalu.
// Po podpieciu prawdziwych czujnikow warto go wlaczyc - wtedy
// martwy czujnik nie zatrzyma proby, tylko zglosi sie sam przez
// xStepTimeout i licznik nTimeouts.
//
// Kroki konczone czujnikiem:
//   st.2 -> st.3    IN2      st.7 -> st.8    IN7
//   st.3 -> st.4    IN3/IN4  st.8 -> st.11   IN8
//   st.6 -> st.7    IN5      st.12-> st.13   IN6
//   st.15-> st.16   IN10
//
// STACJA 1 nie ma czujnika w tej probie. Zamiast niego dziala
// bit xSt01_StackReady: TRUE = stoi tam stos i mozna nim jechac,
// zbocze 0 -> 1 = przyjechal nowy stos (licznik nStacksSeen).
//
// STACJA 4 bada JADACA palete - patrz ACT_MoveSt04.
//
// Wyjatkiem jest przejazd poprzeczny 8 -> 10: tam paleta lezy
// na lancuchu, rolki stacji 8 i 10 sa opuszczone i MUSZA stac.
// Jedzie sam falownik 7, przez tChainTime.
//
// -------------------------------------------------------------
// CO NIE JEST URUCHAMIANE
// -------------------------------------------------------------
// Falowniki 1, 2 i 3 sa ZABLOKOWANE w axDriveEnabled:
//   1  krzywka desztaplarki   - mechanika niegotowa
//   2  krzywka na stacji 8    - mechanika niegotowa
//   3  rolki dociskowe st. 4  - to nie jest transporter
//
// Blokada dziala niezaleznie od tabeli krokow: nawet gdyby
// krok zazadal takiego napedu, nie ruszy. Zeby go dopuscic,
// trzeba swiadomie ustawic bit w axDriveEnabled.
//
// -------------------------------------------------------------
// STEROWANIE
// -------------------------------------------------------------
//   START_TEST = TRUE   symulacja ruchu jedzie
//   START_TEST = FALSE  wszystkie napedy staja
//
//   xCmdResetDrives     kasuje bledy wszystkich falownikow,
//                       dziala na zbocze i sam sie zdejmuje
//
// Po wcisnieciu START maszyna sama sprawdza, czy ktorys naped
// nie stoi w bledzie, i probuje go skasowac - zanim cokolwiek
// ruszy. Jesli sie nie uda, zapala sie xResetFailed.
//
// Pelna aplikacja siedzi w PRG_Machine i na razie nie jest
// wywolywana.
VAR

	// =========================================================
	// STEROWANIE
	// =========================================================

	// GLOWNY BIT TESTU TRASY. TRUE = jedziemy, FALSE = stop.
	START_TEST			: BOOL;


	// =========================================================
	// PROBA CALOSCIOWA: DOWOZ -> DESZTAPLOWANIE -> STACJA 4
	// =========================================================
	//
	// Niezalezna od START_TEST. Wozi palety ze stacji 1 do
	// desztaplarki, potem kazda zwolniona palete przez stacje 4
	// z testem dociskow i ZATRZYMUJE ja na koncu stacji 4.
	// Palete zabiera sie stamtad recznie.

	// Potwierdzenie operatora: palety leza na stacji 1.
	// Kod sam go zdejmuje po przyjeciu - kolejny stos wymaga
	// podania go od nowa.
	xSt01_StackReady	: BOOL;

	// Start dowozu i obslugi transportu w tej probie
	START_FEED			: BOOL;

	// Ile palet przeszlo przez stacje 4
	nFeedPallets		: UDINT;

	// Podglad
	nFeedStep			: INT;
	sFeedPhase			: STRING(79);

	// Wewnetrzne sekwencji dowozu
	nFeedStepOld		: INT;
	xFeedNewStep		: BOOL;
	xFeedArmed			: BOOL;
	xFeedAdvance		: BOOL;
	tFeedStep			: TIME;
	tonFeedStep			: TON;
	rtrgFeedStart		: R_TRIG;

	// =========================================================
	// TOR WYJSCIOWY - DRUGA PALETA W MASZYNIE
	// =========================================================
	//
	// Transport jest rozbity na DWA niezalezne tory:
	//
	//   nFeedStep  tor A: stacja 1 -> 3 -> 4 -> cykl stacji 5
	//   nOutStep   tor B: stacja 5 -> 6 -> ... -> 16
	//
	// Dzieki temu paleta po rozrywaniu jedzie w strone stacji 16
	// SAMA, a desztaplarka moze w tym czasie wydac nastepna.
	// W maszynie sa wtedy dwie palety naraz.
	//
	// Zasob wspolny to transporter stacji 5 (naped 5) i blokada.
	// Dlatego tor A nie wjedzie na stacje 5, dopoki tor B z niej
	// nie zjedzie - patrz krok 75.
	//
	// nOutStep = 0 znaczy TOR B WOLNY.

	nOutStep			: INT;
	sOutPhase			: STRING(79);

	nOutStepOld			: INT;
	xOutNewStep			: BOOL;
	xOutArmed			: BOOL;
	xOutAdvance			: BOOL;
	tOutStep			: TIME;
	tonOutStep			: TON;

	// Stacja 5 skonczyla cykl i oddala palete torowi B.
	// Na tym sygnale desztaplarka wypuszcza nastepna palete.
	xSt05_Done			: BOOL;

	// Zadania startu torow. Tor URUCHAMIA SIE SAM, w swoim kroku 0.
	// Powod jest w komentarzu przy silniku krokow nizej - w skrocie:
	// krok wpisany z ZEWNATRZ wykonalby sie jeszcze w tym samym
	// cyklu, ze stara flaga xOutAdvance, i przeskoczylby natychmiast.
	// -----------------------------------------------------
	// STACJA 8 - POSADZENIE PALETY NOK NA LANCUCHU
	// -----------------------------------------------------
	//
	// Na stacji 8 nie ma blokady, a transporter chodzi tak
	// gladko, ze paleta zatrzymuje sie raz dalej, raz blizej.
	// Dlatego po tSt08_DropDelay od IN7 OPUSZCZAMY rolki: paleta
	// siada na lancuchu i to on ja wyhamowuje - zawsze tak samo.
	//
	// DOTYCZY WYLACZNIE PALET NOK, bo tylko one jada lancuchem.
	// Paleta OK jedzie dalej rolkami i zatrzymuje sie jak dotad -
	// dla niej nic sie nie zmienia.
	//
	// Dwie NIEZALEZNE czasowki od tego samego IN7:
	//   tFeedSt08Stop   zdjecie zadania z falownika (dobieg)
	//   tSt08_DropDelay opuszczenie rolek pod paleta
	tSt08_DropDelay		: TIME := T#830MS;
	tonSt08Drop			: TON;

	// Zatrzask: rolki stacji 8 maja zostac w dole, dopoki lancuch
	// nie zabierze palety. Bez niego kroki, ktore ich nie pisza,
	// podnosilyby je z powrotem.
	xSt08_RollDown		: BOOL;

	// Paleta jest na stacji 8 - od potwierdzenia IN7 do zabrania
	// jej przez lancuch. Na tej fladze chodzi tonSt08Drop, dzieki
	// czemu odliczanie NIE ZALEZY od tego, w ktorym kroku toru B2
	// paleta akurat stoi.
	xSt08_AtStation		: BOOL;

	// Czy TA paleta jedzie trasa odrzutu (lancuchem).
	// W tej probie wszystkie palety jada na stacje 16, wiec bit
	// jest TRUE. Gdy dojdzie klasyfikacja OK/NOK, ma go ustawiac
	// wynik badania, a nie operator.
	xSt08_PalletNOK		: BOOL := TRUE;

	xOutStart			: BOOL;
	xOut2Start			: BOOL;
	xOut3Start			: BOOL;

	// Droga ze stacji 5 wolna: tor B1 pusty i stacja 7 pusta
	xSt05_CanPass		: BOOL;

	// -----------------------------------------------------
	// BUFOROWANIE - TOR B ROZBITY NA TRZY ODCINKI
	// -----------------------------------------------------
	//
	// Odcinki wyznaczaja CZUJNIKI, bo tylko one wiedza, gdzie
	// naprawde stoi paleta:
	//
	//   nOutStep   B1  st.5 -> 6 -> 7    konczy sie na IN5
	//   nOut2Step  B2  st.7 -> 8         konczy sie na IN7
	//   nOut3Step  B3  st.8 -> ... -> 16 konczy sie na IN10
	//
	// Kazdy odcinek zwalnia sie DOPIERO wtedy, gdy nastepny
	// przejmie palete. Dzieki temu w obiegu moga byc naraz:
	// paleta na stacji 5, paleta na 7, paleta na 8 i paleta
	// w drodze na 16 - zamiast jednej na cala maszyne.
	//
	// Transporter stacji 7 (naped 11) obsluguje B1 i B2, a rolki
	// stacji 8 (naped 12) B2. Dlatego paleta czeka w krokach
	// 205 i 218 z ZATRZYMANYMI napedami, zamiast dojezdzac
	// wprost na zajety odcinek.

	nOut2Step			: INT;
	sOut2Phase			: STRING(79);
	nOut2StepOld		: INT;
	xOut2NewStep		: BOOL;
	xOut2Armed			: BOOL;
	xOut2Advance		: BOOL;
	tOut2Step			: TIME;
	tonOut2Step			: TON;

	nOut3Step			: INT;
	sOut3Phase			: STRING(79);
	nOut3StepOld		: INT;
	xOut3NewStep		: BOOL;
	xOut3Armed			: BOOL;
	xOut3Advance		: BOOL;
	tOut3Step			: TIME;
	tonOut3Step			: TON;

	// -----------------------------------------------------
	// STACJA 5 - CZAS PCHANIA PALETY DO BLOKADY
	// -----------------------------------------------------
	//
	// Paleta opiera sie o blokade duzo wczesniej, niz konczy sie
	// krok 80. Kazda sekunda ponad to jest transporterem
	// mielacym pod stojaca paleta - tak przeciazamy naped 5.
	// Po tym czasie napedy 4 i 5 STAJA, a krok trwa dalej.
	//
	// DOMYSLNIE ROWNE tFeedToSt05 - czyli tak, jak bylo przed
	// wprowadzeniem tej nastawy. Moje 4 s bylo za krotkie
	// i paleta nie dojezdzala do blokady.
	//
	// Skracaj DOPIERO po obejrzeniu, gdzie paleta sie zatrzymuje:
	// ma byc na tyle dlugie, zeby doszla do blokady, i na tyle
	// krotkie, zeby transporter nie mielil pod nia bez potrzeby.
	tSt05_Push			: TIME := T#9S;
	tonSt05Push			: TON;

	// -----------------------------------------------------
	// STACJA 4 - ROLKI DOCISKOWE (NAPED 3)
	// -----------------------------------------------------
	//
	// Kreca sie razem z transporterem stacji 4 (naped 4).
	// Bit ponizej wybiera kierunek obrotu - do ustawienia
	// online, bez pobierania projektu.
	xSt04_RollRev		: BOOL := TRUE;

	// Stan dociskow stacji 4 w tej probie - przepisywany co cykl
	xFeedPressOn		: BOOL;
	xFeedPressLoOn		: BOOL;

	// Czas przejazdu st.4 -> st.5. Stacja 5 nie ma czujnika,
	// wiec dojazd konczy sie czasowka. Dobrane na maszynie.
	tFeedToSt05			: TIME := T#9S;

	// DOBIEG NA STACJI 3. Czujnik IN2 widzi krawedz natarcia
	// stosu, a szczeki maja trafic pod DRUGA palete od dolu -
	// stos musi wiec dojechac jeszcze kawalek po wykryciu.
	//
	// ZERO = stop natychmiast po czujniku, czyli tak, jak bylo.
	// Odpowiednik tSt04_StopDelay dla stacji 4.
	tFeedSt03Stop		: TIME := T#0S;

	// Odstep od zatrzymania palety na stacji 5 do ruszenia
	// mechaniki. Stacja 5 nie ma czujnika, wiec nie wiemy, kiedy
	// paleta oprze sie o blokade - dajemy jej na to czas.
	tSt05_Settle		: TIME := T#8S;

	// Stan mechaniki stacji 5 w tej probie - kazdy krok podaje
	// swoj pelny stan, cewki przepisujemy co cykl.
	xFeed05_Block		: BOOL;		// blokada wysunieta
	xFeed05_Lift		: BOOL;		// szczeki podniesione
	xFeed05_Jaws		: BOOL;		// szczeki zamkniete
	xFeed05_Pull		: BOOL;		// silowniki rozrywajace w gorze

	// Diagnostyka napedow zadanych przez biezacy krok
	nFeedBadDrv			: INT;
	sFeedDrvWhy			: STRING(31);
	tonFeedDrv			: TON;

	// -----------------------------------------------------
	// CZASOWKI PRZEJAZDOW BEZ CZUJNIKA
	// -----------------------------------------------------
	//
	// Odcinki, na ktorych nie ma czym potwierdzic dojazdu.
	// Tam, gdzie czujnik jest, czasowka nie jest uzywana wcale.

	tFeed5to6			: TIME := T#12S;		// st.5 -> st.6
	tFeed9Chain			: TIME := T#19S;		// lancuch st.8 -> st.10
	tFeed10to14			: TIME := T#8S;		// st.10 -> st.14
	tFeed14to15			: TIME := T#8S;		// st.14 -> st.15

	// Paleta zniknela z czujnika stacji 16. Po tym czasie
	// uznajemy stacje za pusta - odbiera ja operator.
	tSt16_Clear			: TIME := T#4S;

	// -----------------------------------------------------
	// DOBIEGI PO CZUJNIKACH
	// -----------------------------------------------------
	//
	// Czujnik widzi krawedz natarcia palety, a ona ma stanac
	// na srodku stacji. ZERO = stop natychmiast po czujniku.
	// Odpowiedniki tFeedSt03Stop i tSt04_StopDelay.

	tFeedSt08Stop		: TIME := T#740MS;		// IN7  stacja 8
	tFeedSt16Stop		: TIME := T#0S;		// IN10 stacja 16

	// Rolki podnoszone stacji 8 i 10. TRUE = w gorze, czyli
	// transport wzdluz. Na czas przejazdu lancuchem OBIE musza
	// zejsc, inaczej szarpalyby palete z dwoch stron.
	xFeedRoll08Up		: BOOL := TRUE;
	xFeedRoll10Up		: BOOL := TRUE;

	// Zezwolenie z lancucha bezpieczenstwa
	xSafetyOK			: BOOL := TRUE;

	// KASOWANIE BLEDOW WSZYSTKICH FALOWNIKOW - dziala na zbocze.
	// Bit sam sie zdejmuje po wystawieniu impulsu.
	xCmdResetDrives		: BOOL;

	// Automatyczne kasowanie bledow po wcisnieciu START.
	// FALSE = start nie probuje niczego kasowac.
	xAutoResetOnStart	: BOOL := TRUE;

	// Odstep miedzy kolejnymi probami kasowania
	tResetGap			: TIME := T#1S;

	// Czestotliwosc BAZOWA transporterow [Hz]. Uzywana wszedzie,
	// gdzie alrDriveFreq nie ma wpisanej wlasnej wartosci.
	lrTestFreq			: LREAL := 20.0;

	// =========================================================
	// CZESTOTLIWOSC OSOBNO DLA KAZDEGO NAPEDU [Hz]
	// =========================================================
	//
	// Zero znaczy "uzyj lrTestFreq". Wpisanie liczby dotyczy
	// tylko tego jednego falownika.
	//
	// Przydzial stacja -> falownik:
	//   st.1  -> 8     st.5  -> 5     st.9  -> 7      st.13 -> 15
	//   st.2  -> 9     st.6  -> 6     st.10 -> 16     st.14 -> 17
	//   st.3  -> 10    st.7  -> 11    st.11 -> 13     st.15 -> 18
	//   st.4  -> 4     st.8  -> 12    st.12 -> 14     st.16 -> 19
	//
	// Krzywki 1 i 2 maja wlasna lrCamFreq i ta tablica ich nie
	// dotyczy.
	//
	// UWAGA: naped czyta czestotliwosc przy STARCIE (M_Start jest
	// wolane na zboczu). Zmiana w trakcie jazdy zadziala dopiero
	// przy nastepnym ruszeniu.

	alrDriveFreq		: ARRAY[1..20] OF LREAL;

	// Czas jednego kroku - przejazd palety miedzy stacjami
	tStepTime			: TIME := T#5S;

	// Przejazd poprzeczny transporterem lancuchowym jest dluzszy
	tChainTime			: TIME := T#6S;

	// Czas jednego ruchu silownika. Czujnikow polozenia jeszcze
	// nie ma, wiec po tym czasie uznajemy ruch za wykonany.
	tCylTime			: TIME := T#2S;

	// Stacja 4 - dociski gorne i dolne maja isc praktycznie razem.
	// Gorne schodza pierwsze, dolne po tym krotkim odstepie,
	// zeby dolne nie uniosly palety. Cofanie jest jednoczesne.
	tSt04_UpToLo		: TIME := T#2200MS;

	// FALSE = same transportery, silowniki stoja
	xCylEnable			: BOOL := TRUE;


	// =========================================================
	// CZUJNIKI
	// =========================================================
	//
	// FALSE = jedziemy na samych czasowkach, tak jak dotad.
	// TRUE  = kroki wypisane w ACT_Move koncza sie czujnikiem,
	//         a czasowka pracuje juz tylko jako watchdog.

	xUseSensors			: BOOL := TRUE;

	// STACJA 1 - czujnika IN1 NIE uzywamy. Zastepuje go bit
	// xSt01_StackReady zadeklarowany na gorze.
	nStacksSeen			: UDINT;

	// Obraz czujnikow sprowadzony do JEDNEGO znaczenia:
	// TRUE = PALETA JEST. Polaryzacje ustawia ACT_Inputs i tylko on.
	xPal_St03			: BOOL;		// IN2   stacja 3
	xPal_St04In			: BOOL;		// IN3   wjazd na stacje 4
	xPal_St04End		: BOOL;		// IN4   koniec testu desek
	xPal_St07			: BOOL;		// IN5   stacja 7
	xPal_St13			: BOOL;		// IN6   koniec stacji 13
	xPal_St08			: BOOL;		// IN7   stacja 8
	xPal_St11			: BOOL;		// IN8   stacja 11
	xPal_St16			: BOOL;		// IN10  stacja 16

	// Surowe wejscia - do podgladu bez otwierania GVL
	axInRaw				: ARRAY[1..10] OF BOOL;

	// -----------------------------------------------------
	// POLARYZACJA CZUJNIKOW - JEDYNE MIEJSCE
	// -----------------------------------------------------
	//
	// TRUE  = czujnik ROZWIERA przy palecie (0 = paleta)
	// FALSE = czujnik ZWIERA przy palecie   (1 = paleta)
	//
	// Wartosci ponizej sa wg opisu z maszyny. Jesli ktorys
	// czujnik zachowa sie odwrotnie, przestawia sie JEDEN bit
	// online - bez zmiany kodu i bez pobierania projektu.
	//
	//   1  st.1              nieuzywany
	//   2  st.3              ROZWIERA - stwierdzone na maszynie,
	//                        wbrew pierwotnemu opisu
	//   3  wjazd st.4        rozwiera
	//   4  koniec testu st.4 rozwiera
	//   5  st.7              zwiera
	//   6  koniec st.13      rozwiera
	//   7  st.8              zwiera
	//   8  st.11             zwiera
	//   9  niepodlaczony
	//  10  st.16             zwiera

	axInInverted		: ARRAY[1..10] OF BOOL :=
	                      [FALSE, TRUE, TRUE, TRUE, FALSE,
	                       TRUE, FALSE, FALSE, FALSE, FALSE];

	// WATCHDOG KROKU CZUJNIKOWEGO.
	//
	// FALSE = krok czeka na czujnik BEZ KONCA. Tak jedziemy przy
	//         recznym wyzwalaniu czujnikow - nic nie przeskoczy
	//         kroku, dopoki sam nie podasz sygnalu.
	// TRUE  = po tMoveTimeout krok konczy sie mimo wszystko,
	//         zapala sie xStepTimeout i rosnie nTimeouts.
	xStepWatchdog		: BOOL := FALSE;

	tMoveTimeout		: TIME := T#20S;
	xStepTimeout		: BOOL;
	nTimeouts			: UDINT;


	// =========================================================
	// STACJA 4 - TEST NA JADACEJ PALECIE
	// =========================================================
	//
	// Paleta nie zatrzymuje sie pod rolkami. Czujnik wjazdu (IN3)
	// odlicza tSt04_EntryToPress i wtedy rolki schodza na deski.
	// Czujnik konca testu (IN4) NATYCHMIAST je cofa, a transporter
	// stoi tSt04_StopDelay pozniej - paleta dojezdza do konca stacji.

	tSt04_EntryToPress	: TIME := T#2600MS;
	tSt04_StopDelay		: TIME := T#300MS;


	// =========================================================
	// SZTAPLARKA I DESZTAPLARKA
	// =========================================================
	//
	// Dwa NIEZALEZNE cykle, kazdy z wlasnym bitem startu. Nie
	// maja nic wspolnego z START_TEST.
	//
	// Poziom TRUE = cykl pracuje.
	// Poziom FALSE = natychmiastowy stop, hamulec zaklada sie
	//                tCamBrakeHold pozniej.
	//
	// REGULA NADRZEDNA obu maszyn: nic w szczekach = szczeki
	// OTWARTE i jazda na pozycje DOLNA, niezaleznie od tego,
	// gdzie wozek stoi. Cykl zaczyna sie i konczy na dole
	// z otwartymi szczekami.

	START_DESTACK		: BOOL;		// desztaplarka, stacja 3
	START_STACK			: BOOL;		// sztaplarka, stacja 11

	// -----------------------------------------------------
	// JAZDA RECZNA KRZYWKA
	// -----------------------------------------------------
	//
	// Trzymasz bit - wozek jedzie. Puszczasz - staje, hamulec
	// zaklada sie tCamBrakeHold pozniej, tak samo jak w cyklu.
	//
	// Dziala TYLKO przy zdjetym starcie danej maszyny, zeby
	// nigdy nie walczyc z sekwencja. Sluzy do sprawdzenia,
	// czy enkoder liczy i w ktora strone.

	JOG_DESTACK_FWD		: BOOL;
	JOG_DESTACK_REV		: BOOL;
	JOG_STACK_FWD		: BOOL;
	JOG_STACK_REV		: BOOL;

	xDeJog				: BOOL;
	xStJog				: BOOL;

	// -----------------------------------------------------
	// UCZENIE POZYCJI
	// -----------------------------------------------------
	//
	// Dojedz jogiem tam, gdzie wozek ma stawac, i podaj bit.
	// Zbocze 0 -> 1 przepisuje BIEZACA pozycje enkodera do
	// odpowiedniej nastawy. Koniec z wpisywaniem liczb z palca.
	//
	// UWAGA: nastawy siedza na razie w MAIN, wiec pobranie
	// projektu je kasuje. Po ustaleniu przenosimy do GVL_PERSIST.

	TEACH_DE_BOTTOM		: BOOL;
	TEACH_DE_MIDDLE		: BOOL;
	TEACH_DE_TOP		: BOOL;
	TEACH_ST_BOTTOM		: BOOL;
	TEACH_ST_MIDDLE		: BOOL;
	TEACH_ST_TOP		: BOOL;

	rtrgTeach			: ARRAY[1..6] OF R_TRIG;

	// Ostatnio nauczona pozycja - potwierdzenie na podgladzie
	sTeachLast			: STRING(79);

	// Czestotliwosc krzywek. Osobno od transporterow.
	// Nizej niz transportery - wolniej znaczy krotszy dojazd
	// po zdjeciu zadania, a wiec mniejszy blad pozycji.
	lrCamFreq			: LREAL := 15.0;

	// Ruch szczek - czujnikow polozenia nie ma
	tJawTime			: TIME := T#2S;


	// Odstep od ZALOZENIA hamulca do chwytu szczekami.
	// Wozek musi sie uspokoic, zanim szczeki wejda pod palete.
	tDeGripDelay		: TIME := T#1S;

	// -----------------------------------------------------
	// POZYCJE I LICZNIKI SIEDZA W GVL_PERSIST
	// -----------------------------------------------------
	//
	// Nastawy:  GVL_PERSIST.St03.Cfg.diPosBottom / Middle / Top
	//           GVL_PERSIST.St11.Cfg.diPosBottom / Middle / Top
	//           GVL_PERSIST.St03.Cfg.nStackSize
	// Liczniki: GVL_PERSIST.St03.Mem.nRemaining / nHeld
	//           GVL_PERSIST.St11.Mem.nHeld
	//
	// Sa NIEULOTNE, wiec przezywaja zanik zasilania, aktywacje
	// konfiguracji i reset cold. Uczenie pozycji zapisuje wprost
	// tam - nie ma drugiej kopii, ktora moglaby sie rozjechac.



	// Wyprzedzenie hamowania - zadanie znika tyle przed celem.
	// Zaczynamy od zera i ustawiamy z odczytu diCoast.
	diCamStopLead		: DINT := 0;

	// Okno "jestem na miejscu" przy bazowaniu. Bez niego wozek
	// stojacy tuz przy dolnej pozycji robilby caly obrot, zeby
	// do niej "dojechac".
	diCamTol			: DINT := 300;

	// Ile impulsow za celem uznajemy jeszcze za "jestem".
	// Musi byc WIEKSZE niz dojazd po zdjeciu zadania, inaczej
	// wozek stojacy tuz ZA punktem objechalby caly obrot,
	// zeby do niego wrocic.
	diCamOvershoot		: DINT := 5000;

	// -----------------------------------------------------
	// DOKAD JEDZIE BIEZACY KROK
	// -----------------------------------------------------
	//
	// Krok podaje WARTOSC ENKODERA, do ktorej ma dojechac,
	// a droge liczymy raz, przy wejsciu w krok, z zywej
	// pozycji. Nigdzie nie zakladamy, ile impulsow ma cykl
	// maszyny - to bylo zrodlo kumulujacego sie bledu.

	diDeGoToEnc			: DINT;
	diStGoToEnc			: DINT;

	// -----------------------------------------------------
	// POMIAR - ILE IMPULSOW MA NAPRAWDE CYKL MASZYNY
	// -----------------------------------------------------
	//
	// diDeCycleCounts   droga przejechana miedzy kolejnymi
	//                   dolnymi pozycjami. Jesli enkoder jest
	//                   1:1 z korba, ma byc okolo 65536.
	//                   Kazda inna liczba znaczy, ze cykl
	//                   maszyny to nie jest jeden obrot enkodera.
	// diDeBottomErr     o ile minelismy nauczony dol, ze znakiem
	// diDeCoastMax      najwiekszy zaobserwowany dojazd. Musi
	//                   byc MNIEJSZY niz diCamOvershoot, inaczej
	//                   ruch do punktu tuz za nami pojedzie
	//                   dookola.

	diDeCycleCounts		: DINT;
	diDeBottomErr		: DINT;
	diDeCoastMax		: DINT;

	diStCycleCounts		: DINT;
	diStBottomErr		: DINT;
	diStCoastMax		: DINT;

	// Ustawienie punktu odniesienia osi, impuls jednocyklowy
	xDeSetAccum			: BOOL;
	xStSetAccum			: BOOL;
	diDeAccumSet		: DINT;
	diStAccumSet		: DINT;

	// Roboczy
	diTmp				: DINT;

	// -----------------------------------------------------
	// KONTROLA POPRAWNOSCI NASTAW POZYCJI
	// -----------------------------------------------------
	//
	// Trzy pozycje musza byc od siebie ODDALONE. Zerowe albo
	// pomylone nastawy oznaczaja, ze wozek "juz jest na miejscu"
	// w kazdym kroku - a wtedy szczeki zamykaja sie na dole,
	// na stosie. Cykl nie ma prawa ruszyc na takich nastawach.

	xDeCfgOK			: BOOL;
	xStCfgOK			: BOOL;
	diCamMinSpan		: DINT := 1000;

	// -----------------------------------------------------
	// KONTROLA ENKODERA PO STARCIE
	// -----------------------------------------------------
	//
	// Enkoder absolutny powinien utrzymac wartosc przez zanik
	// zasilania. Zapamietujemy ja na biezaco w GVL_PERSIST
	// i po starcie porownujemy z odczytem. Zgadza sie -
	// bazowanie jest zbedne. Nie zgadza sie - kod to zglasza,
	// zamiast po cichu jechac wedlug zlych pozycji.

	xEncCheckDone		: BOOL;
	diDeEncJump			: DINT;
	diStEncJump			: DINT;
	sEncCheck			: STRING(79);

	// Ile impulsow roznicy jeszcze wybaczamy po starcie
	diEncCheckTol		: DINT := 500;

	// START: wyprzedzenie zdjecia hamulca przed komenda dla
	// falownika. ZERO = jednoczesnie, i tak ma byc.
	tCamBrakeRelease	: TIME := T#0S;

	// STOP: ile hamulec czeka po zdjeciu komendy z falownika.
	// Rampa hamowania falownika to 1 s, wiec hamulec zaciska sie
	// na wolno obracajacym sie jeszcze wale - SWIADOMIE, zeby
	// nie puszczac wozka wolno.
	tCamBrakeHold		: TIME := T#700MS;

	// Kasowanie czuwaka obu osi, dziala na zbocze
	RESET_CAM			: BOOL;

	// =========================================================
	// RESET CYKLU DO ZERA
	// =========================================================
	//
	// Po recznym oproznieniu maszyny z palet. Sprowadza obie
	// maszyny i transport do kroku 0, zeruje liczniki palet
	// i uzgodnienia, kasuje czuwaki osi.
	//
	// NICZYM NIE RUSZA. Wozki wroca na dol dopiero przy starcie,
	// bo krok 0 obu maszyn to "szczeki otwarte, jazda na dol".
	//
	// Bit sam sie zdejmuje.

	RESET_CYCLE			: BOOL;
	rtrgResetCycle		: R_TRIG;

	// -----------------------------------------------------
	// PODGLAD OSI
	// -----------------------------------------------------

	fbCamDestack		: FB_CamAxis;
	fbCamStack			: FB_CamAxis;

	nDeStep				: INT;
	nStStep				: INT;
	sDePhase			: STRING(79);
	sStPhase			: STRING(79);
	nDeCycles			: UDINT;
	nStCycles			: UDINT;

	// -----------------------------------------------------
	// LICZNIKI PALET
	// -----------------------------------------------------
	//
	// GVL_PERSIST.St03.Mem.nRemaining  ile palet zostalo w desztaplarce razem:
	//               na transporterze plus wiszace na szczekach
	// GVL_PERSIST.St03.Mem.nHeld       ile wisi na szczekach desztaplarki
	// GVL_PERSIST.St11.Mem.nHeld       ile palet liczy stos w sztaplarce


	// -----------------------------------------------------
	// UZGODNIENIA Z TRANSPORTEM
	// -----------------------------------------------------

	// Desztaplarka zwolnila palete - transport moze ja zabrac
	xDe_PalletReleased	: BOOL;

	// Desztaplarka pusta, cykl zamkniety na pozycji dolnej
	xDe_Empty			: BOOL;

	// Sztaplarka ma pelny stos na transporterze
	xSt_StackReady		: BOOL;

	// -----------------------------------------------------
	// CZASOWKI OD ZALOZENIA HAMULCA
	// -----------------------------------------------------
	//
	// Licza dopiero od chwili, w ktorej hamulec sie ZACISNIE -
	// nie od wejscia w krok.

	tonDeBrake			: TON;
	tonStBrake			: TON;
	tDeBrakeWait		: TIME;
	tStBrakeWait		: TIME;

	// Czujnik musi byc najpierw WOLNY, zeby sie zaliczyl
	xDeArmed			: BOOL;
	xStArmed			: BOOL;

	// Stan szczek deklarowany przez KAZDY krok i przepisywany
	// na cewki co cykl. Poleganie na tym, ze cewka zachowa
	// wartosc miedzy krokami, juz raz nas kosztowalo prawdziwy
	// blad - ACT_ClearCoils zeruje je w kazdym cyklu.
	xDeJawsClosed		: BOOL;
	xStJawsClosed		: BOOL;

	// -----------------------------------------------------
	// ZYCIE ENKODEROW
	// -----------------------------------------------------
	//
	// Rosna przy KAZDEJ zmianie pozycji. Jesli silnik chodzi,
	// a licznik stoi - enkoder nie jest podlinkowany albo nie
	// liczy. To rozstrzyga sprawe w jednej liczbie.

	nDeEncMoves			: UDINT;
	nStEncMoves			: UDINT;
	diDePosOld			: DINT;
	diStPosOld			: DINT;

	tonDeStep			: TON;
	tonStStep			: TON;
	xDeAdvance			: BOOL;
	xStAdvance			: BOOL;
	tDeStep				: TIME;
	tStStep				: TIME;

	// Zadanie dla osi - liczone przez maszyne stanow,
	// podawane do bloku JEDNYM wywolaniem na cykl
	xDeGo				: BOOL;
	xStGo				: BOOL;
	diDeTarget			: DINT;
	diStTarget			: DINT;

	// Wykrycie zmiany kroku. Bez tego krok zaliczylby xInPos
	// z POPRZEDNIEJ pozycji i przeskoczyl dwa kroki naraz.
	nDeStepOld			: INT;
	nStStepOld			: INT;
	xDeNewStep			: BOOL;
	xStNewStep			: BOOL;
	xDeAtPos			: BOOL;
	xStAtPos			: BOOL;

	rtrgDeStart			: R_TRIG;
	rtrgStStart			: R_TRIG;

	// Cewki hamulcow. TRUE = hamulec ROZLACZONY.
	xBrakeDestack		: BOOL;
	xBrakeStack			: BOOL;


	// =========================================================
	// RECZNE STEROWANIE POJEDYNCZYM SILOWNIKIEM
	// =========================================================
	//
	// Do sprawdzenia okablowania bez sekwencji. Gdy nManCyl <> 0,
	// sekwencja stoi, transportery stoja, a wybrany silownik
	// slucha bitow ponizej.
	//
	//    1  st.3  szczeki desztaplarki
	//    2  st.4  dociski gorne
	//    3  st.4  dociski dolne
	//    4  st.5  blokada
	//    5  st.5  podnoszenie szczek
	//    6  st.5  szczeki (zamkniecie / otwarcie)
	//    7..12 st.5 silowniki rozrywajace 1..6
	//   13  st.8  rolki podnoszone
	//   14  st.10 rolki podnoszone
	//   15  st.11 szczeki sztaplarki

	nManCyl				: INT;
	xManExtend			: BOOL;
	xManRetract			: BOOL;


	// =========================================================
	// DOPUSZCZENIE NAPEDOW
	// =========================================================
	//
	// FALSE = naped nie ruszy, chocby krok tego zadal.
	// Ustawiane w ACT_Config, mozna zmieniac online.

	axDriveEnabled		: ARRAY[1..20] OF BOOL;


	// =========================================================
	// KIERUNEK OBROTOW
	// =========================================================
	//
	// TRUE = jazda w druga strone. Silniki stacji 1, 5, 6, 7,
	// 8, 9, 14, 15, 16 sa podlaczone odwrotnie - do poprawy
	// w szafie, na razie odwracamy bit.

	axReverse			: ARRAY[1..20] OF BOOL;


	// =========================================================
	// PODGLAD
	// =========================================================

	// Gdzie jest wirtualna paleta i co sie z nia dzieje
	nIdx				: INT;		// pozycja na trasie
	nSub				: INT;		// krok sekwencji stacji
	xMoving				: BOOL;		// TRUE = przejazd, FALSE = praca stacji
	sPhase				: STRING(79);

	// Ktore napedy maja teraz pracowac
	axRunReq			: ARRAY[1..20] OF BOOL;

	// Stan napedow
	aeDrvState			: ARRAY[1..20] OF E_NordSK550P_State;
	axDrvRunning		: ARRAY[1..20] OF BOOL;
	alrDrvFreqAct		: ARRAY[1..20] OF LREAL;

	// UWAGA - to sa DWIE ROZNE rzeczy:
	//   axDrvFault  blad zglaszany przez falownik (bit 3 StatusWord)
	//   axDrvError  jakakolwiek blokada: blad, brak zezwolenia
	//               albo zerwana komunikacja
	axDrvFault			: ARRAY[1..20] OF BOOL;
	axDrvError			: ARRAY[1..20] OF BOOL;

	// Slowa sterujace i statusowe - do czytania, co naped
	// naprawde zglasza
	awDrvStatus			: ARRAY[1..20] OF UINT;
	awDrvControl		: ARRAY[1..20] OF UINT;

	// Ktorykolwiek naped zglasza blad
	xAnyDriveError		: BOOL;
	xAnyDriveFault		: BOOL;

	// Kasowanie nie poskutkowalo - blad wraca albo trzyma
	xResetFailed		: BOOL;

	// Trwa kasowanie bledow przed startem
	xResetInProgress	: BOOL;
	nResetTries			: INT;

	// Blokada zadzialala - lancuch wymusil postoj rolek 8 i 10
	xChainInterlock		: BOOL;

	// Blokada stacji 5 kontra transporter - patrz ACT_ApplyDrives
	xSt05_BlockLock		: BOOL;
	tonSt05BlockDown	: TON;

	// Czas biezacego kroku
	tThisStep			: TIME;

	// Licznik pelnych przebiegow trasy
	nLoops				: UDINT;

	// =========================================================
	// LICZNIKI ZYCIA - do sprawdzenia, co sie naprawde wykonuje
	// =========================================================
	//
	// nCycles     rosnie w kazdym cyklu zadania. Jesli stoi,
	//             MAIN sie nie wykonuje albo wysypal sie wczesniej.
	// nOutWrites  rosnie za kazdym przepisaniem cewek na wyjscia.
	//             Jesli nCycles rosnie, a nOutWrites stoi -
	//             program nie dochodzi do ACT_Outputs.
	// nCoilsOn    ile cewek jest w tej chwili podanych. Jesli
	//             rosnie i spada, a nic sie nie rusza - sygnal
	//             nie dochodzi do zaworu.

	nCycles				: UDINT;
	nOutWrites			: UDINT;
	nCoilsOn			: INT;


	// =========================================================
	// CEWKI ZAWOROW
	// =========================================================
	//
	// Stan trzymany miedzy cyklami. ACT_Outputs przepisuje go
	// na wyjscia - mapowanie jest TAM i tylko tam.

	// Stacja 3 - szczeki desztaplarki
	xSt03_JawClose		: BOOL;
	xSt03_JawOpen		: BOOL;

	// Stacja 4 - dociski. Obie grupy gornych chodza razem.
	xSt04_UpExt			: BOOL;
	xSt04_UpRet			: BOOL;
	xSt04_LoExt			: BOOL;
	xSt04_LoRet			: BOOL;

	// Stacja 5
	xSt05_BlockExt		: BOOL;		// blokada wysuw
	xSt05_BlockRet		: BOOL;		// blokada opuszczenie
	xSt05_LiftUp		: BOOL;		// szczeki w gore
	xSt05_LiftDown		: BOOL;		// szczeki w dol
	xSt05_JawClose		: BOOL;		// trzy pary szczek razem
	axSt05_PullUp		: ARRAY[1..6] OF BOOL;
	axSt05_PullDown		: ARRAY[1..6] OF BOOL;

	// Rolki podnoszone
	xSt08_Up			: BOOL;
	xSt08_Down			: BOOL;
	xSt10_Up			: BOOL;
	xSt10_Down			: BOOL;

	// Stacja 11 - szczeki sztaplarki
	xSt11_JawClose		: BOOL;
	xSt11_JawOpen		: BOOL;


	// =========================================================
	// NAPEDY
	// =========================================================

	fbNord				: ARRAY[1..20] OF FB_NordSK550PP;


	// =========================================================
	// OBSERWATOR STANU - LOG CSV NA DYSKU STEROWNIKA
	// =========================================================
	//
	// Co tLogPeriod jeden wiersz z kluczowymi zmiennymi, a do
	// tego wiersz na kazde ZDARZENIE: zmiana numeru kroku,
	// czujnika, zadania napedu, bledu falownika, bitu operatora,
	// szczek, skok enkodera. Najwyzej jeden wiersz na cykl.
	//
	// Nowy plik: start PLC, RESET_CYCLE, zbocze xLogNewFile.
	// Katalog MUSI istniec na sterowniku: fbLog.sDir
	// (domyslnie C:\TesterPalet\log\). Nazwa pliku w fbLog.sFileName.
	//
	// Logger tylko CZYTA zmienne procesu - ACT_Logger idzie jako
	// ostatnia akcja cyklu, po ACT_Outputs, zeby w pliku bylo to,
	// co naprawde poszlo na wyjscia.

	fbLog				: FB_CsvLogger;

	// FALSE = nie zbieramy wierszy (plik zostaje, nic sie nie psuje)
	xLogEnable			: BOOL := TRUE;

	// Zbocze = nowy plik bez resetu cyklu. Sam sie zdejmuje.
	xLogNewFile			: BOOL;

	// Takt wiersza okresowego
	tLogPeriod			: TIME := T#1S;
	tonLog				: TON;

	// Skok enkodera w jednym cyklu, od ktorego piszemy zdarzenie
	diLogEncJump		: DINT := 2000;

	// Powod biezacego wiersza - do kolumny "why"
	sLogWhy				: STRING(79);
	xLogEvent			: BOOL;
	nLogRows			: UDINT;

	// Pamiec do wykrywania zdarzen
	xLogInit			: BOOL;
	anLogStepOld		: ARRAY[1..6] OF INT;
	axLogInOld			: ARRAY[1..10] OF BOOL;
	axLogReqOld			: ARRAY[1..20] OF BOOL;
	axLogFaultOld		: ARRAY[1..20] OF BOOL;
	axLogBitOld			: ARRAY[1..24] OF BOOL;
	axLogBit			: ARRAY[1..24] OF BOOL;

	// Robocze do skladania nazw kolumn napedow
	sLogPfx				: STRING(15);
	wLogFesto1			: WORD;
	wLogFesto2			: WORD;
	nLogI				: INT;
	nLogJ				: INT;


	// =========================================================
	// WEWNETRZNE
	// =========================================================

	xInit				: BOOL;
	i					: INT;
	lrThisFreq			: LREAL;
	tonStep				: TON;
	tonResetGap			: TON;
	xAdvance			: BOOL;
	rtrgStart			: R_TRIG;
	rtrgResetDrv		: R_TRIG;
	rtrgStack			: R_TRIG;
	xDoResetPulse		: BOOL;
	axRunOld			: ARRAY[1..20] OF BOOL;

	// Krok zglasza tu, ze czeka na czujnik i ktory to czujnik.
	// Kasowane co cykl, ustawiane przez sam krok.
	xWaitSensor			: BOOL;
	xSensorOK			: BOOL;

	// Czujnik musi najpierw byc WOLNY. Bez tego zaliczylby sie
	// stan sprzed kroku albo czujnik zawieszony na stale.
	xStepArmed			: BOOL;

	// Wykrycie zmiany kroku - czasowka i uzbrojenie od zera
	xNewStep			: BOOL;
	nIdxOld				: INT;
	nSubOld				: INT;
	xMovingOld			: BOOL;

	// TRUE = przejazd ma jeszcze kroki wewnetrzne, nIdx zostaje
	xHoldIdx			: BOOL;

END_VAR
VAR CONSTANT

	// P105 falownikow
	cFmax				: LREAL := 50.0;

	// Liczba falownikow zmapowanych w .tsproj
	cNumDrives			: INT := 19;

	// Liczba pozycji na trasie
	cLastIdx			: INT := 16;

	// Ile razy probujemy skasowac blad przed startem
	cResetTries			: INT := 3;

END_VAR

alrDriveFreq[12] := 10;



// =============================================================
// MAIN - TEST RUCHU TRANSPORTEROW
// =============================================================

// Puls zycia - jesli ten licznik stoi, MAIN sie nie wykonuje
nCycles := nCycles + 1;

ACT_Config();

ACT_Inputs();

ACT_Sequence();

// Krzywki chodza NIEZALEZNIE od START_TEST i po ACT_Sequence,
// zeby ich szczeki mialy pierwszenstwo przed sekwencja linii.
ACT_CamCycles();

// Transport proby calosciowej - po krzywkach, zeby jego
// cewki i zadania napedow mialy pierwszenstwo.
ACT_TestFeed();

ACT_ResetDrives();

ACT_ApplyDrives();

ACT_Drives();

ACT_Outputs();

// Obserwator stanu - OSTATNI, zeby logowal to, co poszlo na wyjscia
ACT_Logger();

ACTION ACT_ApplyDrives:
// =============================================================
// ACT_ApplyDrives
// Zadanie ruchu -> metody falownikow
// =============================================================
//
// Metody wolamy NA ZBOCZU. Blok napedu przy blokadzie sam kasuje
// zadanie ruchu i naped nie moze ruszyc sam po ustapieniu
// przyczyny - wolanie M_Start co cykl zepsuloby to zabezpieczenie.

xAnyDriveError := FALSE;


// -------------------------------------------------------------
// BLOKADA: LANCUCH KONTRA ROLKI STACJI 8 I 10
// -------------------------------------------------------------
//
// Gdy jedzie transporter lancuchowy, rolki stacji 8 i 10 sa
// opuszczone i paleta lezy na lancuchu. Krecenie nimi w tym
// czasie szarpaloby palete z dwoch stron naraz.
//
// To nie jest poprawka tabeli krokow, tylko warunek nadrzedny -
// zadziala takze wtedy, gdy ktos pozniej zmieni tabele.

xChainInterlock := FALSE;

IF axRunReq[7] THEN

	IF axRunReq[12] OR axRunReq[16] THEN
		xChainInterlock := TRUE;
	END_IF

	axRunReq[12] := FALSE;		// rolki stacji 8
	axRunReq[16] := FALSE;		// rolki stacji 10

END_IF


// -------------------------------------------------------------
// BLOKADA STACJI 5 KONTRA TRANSPORTER
// -------------------------------------------------------------
//
// Wysunieta blokada znaczy "paleta ma tu stanac". Wypychanie jej
// wtedy na stacje 6 to praca transportera w zapore - i to jest
// przyczyna, dla ktorej naped 5 wchodzil w przeciazenie.
//
// WJAZD ZE STACJI 4 JEST WYJATKIEM: tam blokada MA byc wysunieta,
// bo to ona zatrzymuje palete. Dlatego warunek dotyczy wylacznie
// jazdy W STRONE STACJI 6, czyli kroku 180 toru B1.
//
// Blokada nie ma czujnika polozenia, wiec zadamy nie tylko
// zdjetej komendy, ale i tCylTime na jej faktyczne opuszczenie.
// Warunek nadrzedny, jak blokada lancucha wyzej - nie zalezy od
// tabeli krokow i zadziala takze po jej zmianie.

xSt05_BlockLock := FALSE;

IF (nOutStep = 180) AND NOT tonSt05BlockDown.Q THEN
	xSt05_BlockLock := TRUE;
	axRunReq[5] := FALSE;
	axRunReq[6] := FALSE;
END_IF


// -------------------------------------------------------------
// SPRZEZENIE: ROLKI DOCISKOWE STACJI 4 Z TRANSPORTEREM
// -------------------------------------------------------------
//
// Naped 3 (gorne rolki dociskowe) kreci sie zawsze wtedy, gdy
// kreci sie transporter stacji 4 (naped 4). Nie ma sensu, zeby
// rolki lezaly na deskach i staly, kiedy paleta pod nimi jedzie.
//
// Warunek nadrzedny, tak jak blokada lancucha wyzej: nie zalezy
// od tabeli krokow i zadziala takze po jej zmianie.
//
// Kierunek bierzemy z bitu, ktory mozna przestawic online.

axReverse[3] := xSt04_RollRev;

IF axRunReq[4] THEN
	axRunReq[3] := TRUE;
END_IF


FOR i := 1 TO cNumDrives DO

	// Naped niedopuszczony nie ruszy, chocby krok tego zadal
	IF NOT axDriveEnabled[i] THEN
		axRunReq[i] := FALSE;
	END_IF

	IF axDrvError[i] THEN
		xAnyDriveError := TRUE;
	END_IF



	// Czestotliwosc: wlasna dla napedu, inaczej bazowa.
	lrThisFreq := lrTestFreq;

	IF alrDriveFreq[i] > 0.0 THEN
		lrThisFreq := alrDriveFreq[i];
	END_IF

	// Krzywki maja wlasna nastawe i wygrywaja z tablica
	IF (i = 1) OR (i = 2) THEN
		lrThisFreq := lrCamFreq;
	END_IF

	// Naped zablokowany (blad, brak zezwolenia, zerwana
	// komunikacja) SAM kasuje u siebie zadanie ruchu - i slusznie,
	// bo nie wolno mu ruszyc samoczynnie po ustapieniu przyczyny.
	//
	// Warstwa maszyny musi wiec wydac komende OD NOWA. Dlatego:
	//   - w czasie blokady nie wolamy M_Start (byloby bez sensu,
	//     a lamaloby regule wolania na zboczu),
	//   - pamiec zbocza trzymamy wtedy wyzerowana, zeby po
	//     ustapieniu przyczyny powstalo JEDNO nowe zbocze.
	//
	// Bez tego naped, ktory raz wpadl w blad, stalby juz na
	// zawsze - skasowanie bledu nic by nie dalo, bo zbocze
	// startu dawno minelo.

	IF axRunReq[i] AND NOT axRunOld[i] AND NOT axDrvError[i] THEN
		fbNord[i].M_Start(lrFreq := lrThisFreq, xReverse := axReverse[i]);
	END_IF

	IF NOT axRunReq[i] AND axRunOld[i] THEN
		fbNord[i].M_Stop();
	END_IF

	axRunOld[i] := axRunReq[i] AND NOT axDrvError[i];

END_FOR
END_ACTION

ACTION ACT_CamCycles:
// =============================================================
// ACT_CamCycles
// Desztaplarka (st.3) i sztaplarka (st.11)
// =============================================================
//
// KORBA JEDZIE ZAWSZE W JEDNA STRONE. Cykl to jeden obrot:
// dol -> posrednia -> gorna -> DALEJ TYM SAMYM KIERUNKIEM
// z powrotem na dol. Nigdy nie wracamy tam, skad przyjechalismy.
//
// Enkoder jest jednoobrotowy i potrafi pokazac wartosc wieksza
// niz jeden obrot, wiec FB_CamAxis sprowadza ja modulo 65536,
// liczy przyrost ze znakiem i sam wykrywa przejscia przez zero.
// Tutaj operujemy juz tylko pozycjami 0..65535.
//
// REGULA NADRZEDNA obu maszyn: nic w szczekach = szczeki
// OTWARTE i jazda na pozycje DOLNA, niezaleznie od tego, gdzie
// wozek stoi.
//
// -------------------------------------------------------------
// SZCZEKI
// -------------------------------------------------------------
// KAZDY krok deklaruje xDeJawsClosed / xStJawsClosed, a cewki
// przepisujemy raz, na koncu akcji. Nie wolno polegac na tym,
// ze cewka zachowa wartosc miedzy krokami - ACT_ClearCoils
// zeruje wszystkie cewki w kazdym cyklu przy zdjetym START_TEST,
// wiec krok, ktory ich nie odswieza, traci sterowanie zaworem.
//
// -------------------------------------------------------------
// SYGNALY
// -------------------------------------------------------------
//   xPal_St03     IN2   sztapla na stacji 3
//   xPal_St04In   IN3   stacja 4 przyjela palete
//   xPal_St11     IN8   paleta na stacji 11
//
// Czujnik musi byc najpierw WOLNY, zeby sie zaliczyl.


// =============================================================
// RESET CYKLU DO ZERA
// =============================================================
//
// Wykonujemy to PRZED maszynami stanow, zeby jeszcze w tym
// samym cyklu ruszyly juz od kroku 0 - takze transport,
// bo ACT_TestFeed idzie po tej akcji.

rtrgResetCycle(CLK := RESET_CYCLE);

IF rtrgResetCycle.Q THEN

	nDeStep   := 0;
	nStStep   := 0;
	nFeedStep := 0;
	nOutStep  := 0;
	nOut2Step := 0;
	nOut3Step := 0;

	xOutStart  := FALSE;
	xOut2Start := FALSE;
	xOut3Start := FALSE;
	xSt08_RollDown  := FALSE;
	xSt08_AtStation := FALSE;

	xSt05_Done := FALSE;

	GVL_PERSIST.St03.Mem.nRemaining := 0;
	GVL_PERSIST.St03.Mem.nHeld      := 0;
	GVL_PERSIST.St11.Mem.nHeld      := 0;

	xDe_PalletReleased := FALSE;
	xSt_StackReady     := FALSE;
	xSt01_StackReady   := FALSE;

	nFeedPallets := 0;
	nDeCycles    := 0;
	nStCycles    := 0;

	RESET_CYCLE := FALSE;

END_IF


// =============================================================
// KONTROLA NASTAW POZYCJI
// =============================================================
//
// Trzy punkty musza byc od siebie oddalone o co najmniej
// diCamMinSpan, liczac najkrotsza droga po okregu. Zerowe
// nastawy - na przyklad po skasowaniu danych nieulotnych -
// znacza, ze kazdy krok od razu melduje "na pozycji", a szczeki
// zamykaja sie tam, gdzie wozek akurat stoi.

xDeCfgOK := TRUE;

diTmp := GVL_PERSIST.St03.Cfg.diPosMiddle - GVL_PERSIST.St03.Cfg.diPosBottom;
IF diTmp >  32768 THEN diTmp := diTmp - 65536; END_IF
IF diTmp < -32768 THEN diTmp := diTmp + 65536; END_IF
IF ABS(diTmp) < diCamMinSpan THEN xDeCfgOK := FALSE; END_IF

diTmp := GVL_PERSIST.St03.Cfg.diPosTop - GVL_PERSIST.St03.Cfg.diPosBottom;
IF diTmp >  32768 THEN diTmp := diTmp - 65536; END_IF
IF diTmp < -32768 THEN diTmp := diTmp + 65536; END_IF
IF ABS(diTmp) < diCamMinSpan THEN xDeCfgOK := FALSE; END_IF

diTmp := GVL_PERSIST.St03.Cfg.diPosTop - GVL_PERSIST.St03.Cfg.diPosMiddle;
IF diTmp >  32768 THEN diTmp := diTmp - 65536; END_IF
IF diTmp < -32768 THEN diTmp := diTmp + 65536; END_IF
IF ABS(diTmp) < diCamMinSpan THEN xDeCfgOK := FALSE; END_IF


xStCfgOK := TRUE;

diTmp := GVL_PERSIST.St11.Cfg.diPosMiddle - GVL_PERSIST.St11.Cfg.diPosBottom;
IF diTmp >  32768 THEN diTmp := diTmp - 65536; END_IF
IF diTmp < -32768 THEN diTmp := diTmp + 65536; END_IF
IF ABS(diTmp) < diCamMinSpan THEN xStCfgOK := FALSE; END_IF

diTmp := GVL_PERSIST.St11.Cfg.diPosTop - GVL_PERSIST.St11.Cfg.diPosBottom;
IF diTmp >  32768 THEN diTmp := diTmp - 65536; END_IF
IF diTmp < -32768 THEN diTmp := diTmp + 65536; END_IF
IF ABS(diTmp) < diCamMinSpan THEN xStCfgOK := FALSE; END_IF

diTmp := GVL_PERSIST.St11.Cfg.diPosTop - GVL_PERSIST.St11.Cfg.diPosMiddle;
IF diTmp >  32768 THEN diTmp := diTmp - 65536; END_IF
IF diTmp < -32768 THEN diTmp := diTmp + 65536; END_IF
IF ABS(diTmp) < diCamMinSpan THEN xStCfgOK := FALSE; END_IF


// =============================================================
// ZMIANA KROKU
// =============================================================
//
// Blok osi liczy xInPos wzgledem celu z POPRZEDNIEGO cyklu,
// wiec w pierwszym cyklu nowego kroku tej informacji nie
// zaliczamy - inaczej krok przeskoczylby dwa naraz.

// =============================================================
// KONTROLA ENKODERA PO STARCIE
// =============================================================
//
// Raz, w pierwszym cyklu po starcie PLC. Porownujemy odczyt
// z wartoscia zapamietana przed wylaczeniem. Roznica wieksza
// niz diEncCheckTol znaczy, ze enkoder NIE utrzymal pozycji
// i trzeba go zbazowac na dole.

IF NOT xEncCheckDone THEN

	xEncCheckDone := TRUE;

	diTmp := fbCamDestack.diPos - GVL_PERSIST.St03.Mem.diLastPos;
	IF diTmp >  32768 THEN diTmp := diTmp - 65536; END_IF
	IF diTmp < -32768 THEN diTmp := diTmp + 65536; END_IF
	diDeEncJump := diTmp;

	diTmp := fbCamStack.diPos - GVL_PERSIST.St11.Mem.diLastPos;
	IF diTmp >  32768 THEN diTmp := diTmp - 65536; END_IF
	IF diTmp < -32768 THEN diTmp := diTmp + 65536; END_IF
	diStEncJump := diTmp;

	GVL_PERSIST.St03.Mem.xNeedHoming := ABS(diDeEncJump) > diEncCheckTol;
	GVL_PERSIST.St11.Mem.xNeedHoming := ABS(diStEncJump) > diEncCheckTol;

	sEncCheck := 'enkodery utrzymaly pozycje - bazowanie zbedne';

	IF GVL_PERSIST.St03.Mem.xNeedHoming THEN
		sEncCheck := 'DESZTAPLARKA - enkoder nie utrzymal pozycji, zbazuj dol';
	END_IF

	IF GVL_PERSIST.St11.Mem.xNeedHoming THEN
		sEncCheck := 'SZTAPLARKA - enkoder nie utrzymal pozycji, zbazuj dol';
	END_IF

END_IF


// Zapamietanie biezacej pozycji na wypadek zaniku zasilania.
// PLC ma 1 s UPSa, wiec TwinCAT zdazy zapisac dane nieulotne.
GVL_PERSIST.St03.Mem.diLastPos := fbCamDestack.diPos;
GVL_PERSIST.St11.Mem.diLastPos := fbCamStack.diPos;


// Impulsy ustawienia punktu odniesienia - kasowane co cykl
xDeSetAccum := FALSE;
xStSetAccum := FALSE;


xDeNewStep := (nDeStep <> nDeStepOld);
xStNewStep := (nStStep <> nStStepOld);

nDeStepOld := nDeStep;
nStStepOld := nStStep;

IF xDeNewStep THEN
	tonDeStep(IN := FALSE);
	xDeArmed := FALSE;
END_IF

IF xStNewStep THEN
	tonStStep(IN := FALSE);
	xStArmed := FALSE;
END_IF

tonDeStep(IN := TRUE, PT := tDeStep);
tonStStep(IN := TRUE, PT := tStStep);

xDeAdvance := tonDeStep.Q AND NOT xDeNewStep;
xStAdvance := tonStStep.Q AND NOT xStNewStep;

xDeAtPos := fbCamDestack.xInPos AND NOT xDeNewStep;
xStAtPos := fbCamStack.xInPos   AND NOT xStNewStep;


// Czasowki liczone od ZACISNIECIA hamulca, nie od wejscia w krok
tonDeBrake(IN := NOT fbCamDestack.xBrakeRelease, PT := tDeBrakeWait);
tonStBrake(IN := NOT fbCamStack.xBrakeRelease,   PT := tStBrakeWait);


// =============================================================
// DESZTAPLARKA - STACJA 3
// =============================================================
//
//   0   dom: szczeki otwarte, jazda na dol
//   10  czekam na sztaple
//   20  jazda na pozycje posrednia, szczeki OTWARTE
//   30  hamulec zalozony, odliczam 1 s
//   40  szczeki zamykaja sie pod druga paleta od dolu
//   50  jazda na gore - stos uniesiony przez druga palete
//   60  info do transportu, czekam az stacja 4 przyjmie palete
//   70  DALEJ tym samym kierunkiem, dopelnienie obrotu na dol
//   80  hamulec zalozony, szczeki otwieraja sie
//   85  BRAMKA CYKLU - na dole czekam na koniec cyklu stacji 5
//   90  ostatnia paleta - nie ma czego chwytac, wyjezdza sama

xDeJog := (JOG_DESTACK_FWD OR JOG_DESTACK_REV) AND NOT START_DESTACK;

rtrgDeStart(CLK := START_DESTACK);

IF rtrgDeStart.Q THEN
	nDeStep := 0;
END_IF

IF rtrgDeStart.Q AND xAutoResetOnStart AND xAnyDriveFault THEN
	xResetInProgress := TRUE;
	nResetTries      := 0;
	xResetFailed     := FALSE;
END_IF

xDeGo        := FALSE;
tDeStep      := tJawTime;
tDeBrakeWait := tDeGripDelay;


// REGULA NADRZEDNA: pusto w szczekach w kroku niosacym stos
// to sprzecznosc - wracamy do domu zamiast jechac dalej.
IF (GVL_PERSIST.St03.Mem.nHeld <= 0) AND (nDeStep >= 50) AND (nDeStep <= 70) THEN
	nDeStep := 0;
END_IF


IF NOT START_DESTACK THEN
	sDePhase := 'DESZTAPLARKA - stop, START_DESTACK = FALSE';
END_IF

IF xDeJog THEN
	sDePhase := 'DESZT. RECZNIE - jazda krzywka, patrz na diPos';
END_IF

IF START_DESTACK AND fbCamDestack.xBrakeWait THEN
	sDePhase := 'DESZT. czekam na odpuszczenie hamulca przed startem';
END_IF

IF START_DESTACK AND fbCamDestack.xStall THEN
	sDePhase := 'DESZT. CZUWAK - falownik pracuje, a enkoder nie liczy';
END_IF

IF START_DESTACK AND fbCamDestack.xNoDrvAck THEN
	sDePhase := 'DESZT. CZUWAK - falownik 1 nie potwierdza pracy';
END_IF

IF START_DESTACK AND fbCamDestack.xStall AND axDrvFault[1] THEN
	sDePhase := 'DESZT. CZUWAK - falownik 1 w bledzie, kasuj xCmdResetDrives';
END_IF

IF START_DESTACK AND fbCamDestack.xStall AND NOT axDriveEnabled[1] THEN
	sDePhase := 'DESZT. CZUWAK - naped 1 NIEDOPUSZCZONY, ACT_Config sie nie wykonalo';
END_IF


IF START_DESTACK AND NOT xDeCfgOK THEN
	sDePhase := 'DESZT. NASTAWY POZYCJI PUSTE albo BLEDNE - naucz dol/srodek/gore';
END_IF


IF START_DESTACK AND NOT fbCamDestack.xStall AND xDeCfgOK THEN

	CASE nDeStep OF

	0:
		// REGULA NADRZEDNA: nic w szczekach = otwarte i na dol.
		//
		// Szczeki otwieramy OD RAZU, takze na gorze. Swiadomy
		// wybor: przy 1000 Nm na krzywce gorsza awaria jest
		// przeciagniecie zamknietych szczek przez stos niz
		// spadniecie palet. NIE dodawac tu zjazdu "trzymajac"
		// bez rozmowy - bylo zrobione i zostalo cofniete.
		sDePhase := 'DESZT. 0 dom: szczeki otwarte, jazda na dol';
		xDeJawsClosed := FALSE;
		GVL_PERSIST.St03.Mem.nHeld    := 0;
		xDeGo       := TRUE;
		diDeGoToEnc := GVL_PERSIST.St03.Cfg.diPosBottom;
		IF xDeAtPos THEN nDeStep := 10; END_IF

	10:
		sDePhase := 'DESZT. 1 czekam na sztaple na stacji 3 (IN2)';
		xDeJawsClosed := FALSE;
		xDe_Empty := TRUE;

		// Sztapla, ktora JUZ stoi na stacji przy wejsciu w krok,
		// jest sztapla gotowa do pracy - nie kazemy jej zjezdzac
		// i wracac. Uzbrojenie chroni tylko przed policzeniem
		// tej samej sztapli dwa razy w trakcie czekania.
		IF xDeNewStep AND xPal_St03 THEN xDeArmed := TRUE; END_IF

		IF NOT xPal_St03 THEN xDeArmed := TRUE; END_IF

		IF xDeArmed AND xPal_St03 THEN
			GVL_PERSIST.St03.Mem.nRemaining := GVL_PERSIST.St03.Cfg.nStackSize;
			xDe_Empty    := FALSE;
			nDeStep      := 20;
		END_IF

	20:
		sDePhase := 'DESZT. 2 jazda na pozycje posrednia, szczeki otwarte';
		xDeJawsClosed := FALSE;
		xDeGo       := TRUE;
		diDeGoToEnc := GVL_PERSIST.St03.Cfg.diPosMiddle;
		IF xDeAtPos THEN nDeStep := 30; END_IF

	30:
		sDePhase := 'DESZT. 3 hamulec zalozony - odliczam przed chwytem';
		xDeJawsClosed := FALSE;
		IF tonDeBrake.Q THEN nDeStep := 40; END_IF

	40:
		sDePhase := 'DESZT. 4 szczeki chwytaja 2. palete od dolu';
		xDeJawsClosed := TRUE;
		IF xDeAdvance THEN
			GVL_PERSIST.St03.Mem.nHeld := GVL_PERSIST.St03.Mem.nRemaining - 1;
			nDeStep := 50;
		END_IF

	50:
		sDePhase := 'DESZT. 5 jazda na gore - stos uniesiony';
		xDeJawsClosed := TRUE;
		xDeGo       := TRUE;
		diDeGoToEnc := GVL_PERSIST.St03.Cfg.diPosTop;
		IF xDeAtPos THEN nDeStep := 60; END_IF

	60:
		// Potwierdzeniem odbioru jest czujnik na KONCU stacji 4
		// (IN4), a nie ten od wjazdu pod rolki. Dopiero on mowi,
		// ze paleta naprawde zjechala z desztaplarki.
		//
		// TEN WARUNEK MUSI BYC KROTKI. Stos wisi tu na szczekach,
		// wiec nie wolno w tym kroku czekac na nic dalszego niz
		// zjazd palety z desztaplarki - bramka cyklu stoi w
		// kroku 85, na dole, przy stosie opartym o transporter.
		//
		// IN4 pilnuje takze tego, zeby stos nie zjechal na palete,
		// ktora jeszcze nie zdazyla wyjechac.
		sDePhase := 'DESZT. 6 paleta zwolniona - czekam na koniec st.4 (IN4)';
		xDeJawsClosed := TRUE;
		xDe_PalletReleased := TRUE;

		IF NOT xPal_St04End THEN xDeArmed := TRUE; END_IF

		IF xPal_St04End AND NOT xDeArmed THEN
			sDePhase := 'DESZT. 6 IN4 JUZ zaslonony - odslon i zaslon ponownie';
		END_IF

		IF xDeArmed AND xPal_St04End THEN
			GVL_PERSIST.St03.Mem.nRemaining       := GVL_PERSIST.St03.Mem.nRemaining - 1;
			xDe_PalletReleased := FALSE;
			nDeStep            := 70;
		END_IF

	70:
		// DALEJ tym samym kierunkiem - dopelnienie pelnego obrotu
		sDePhase := 'DESZT. 7 dopelnienie obrotu - zjazd stosu na dol';
		xDeJawsClosed := TRUE;
		xDeGo       := TRUE;
		diDeGoToEnc := GVL_PERSIST.St03.Cfg.diPosBottom;
		IF xDeAtPos THEN nDeStep := 80; END_IF

	80:
		sDePhase := 'DESZT. 8 hamulec zalozony - szczeki otwieraja sie';
		tDeBrakeWait := tJawTime;
		GVL_PERSIST.St03.Mem.nHeld := 0;

		xDeJawsClosed := TRUE;

		IF NOT fbCamDestack.xBrakeRelease THEN
			xDeJawsClosed := FALSE;
		END_IF

		IF tonDeBrake.Q AND (GVL_PERSIST.St03.Mem.nRemaining > 1) THEN
			nDeCycles := nDeCycles + 1;
			nDeStep   := 85;
		END_IF

		IF tonDeBrake.Q AND (GVL_PERSIST.St03.Mem.nRemaining = 1) THEN
			nDeCycles := nDeCycles + 1;
			nDeStep   := 90;
		END_IF

		IF tonDeBrake.Q AND (GVL_PERSIST.St03.Mem.nRemaining <= 0) THEN
			nDeStep := 0;
		END_IF

	85:
		// BRAMKA CYKLU - JEDYNE DLUGIE CZEKANIE DESZTAPLARKI.
		//
		// Stoi TU, a nie na gorze w kroku 60, i to jest istota
		// sprawy: wozek jest na dole, stos oparty o transporter,
		// szczeki otwarte, hamulec zalozony. Nic nie wisi.
		//
		// Wczesniej ta bramka stala w kroku 60 i stos zostawal
		// zawieszony na szczekach przez caly cykl stacji 5 -
		// dziesiatki sekund zamiast kilku. Tak stracilismy stos.
		//
		// Czekamy na koniec cyklu stacji 5: dopiero wtedy ma sens
		// wydawac kolejna palete, bo poprzednia zjechala juz
		// w strone stacji 16.
		sDePhase := 'DESZT. 8b stos na dole - czekam na koniec cyklu st.5';
		xDeJawsClosed := FALSE;

		IF xSt05_Done THEN
			xSt05_Done := FALSE;
			nDeStep    := 20;
		END_IF

	90:
		// Ostatnia paleta lezy wprost na transporterze - szczeki
		// nie maja pod co wejsc, wiec wyjezdza sama.
		sDePhase := 'DESZT. 9 ostatnia paleta - wyjezdza sama, bez chwytu';
		xDeJawsClosed := FALSE;
		xDe_PalletReleased := TRUE;

		IF NOT xPal_St04End THEN xDeArmed := TRUE; END_IF

		IF xPal_St04End AND NOT xDeArmed THEN
			sDePhase := 'DESZT. 9 IN4 JUZ zaslonony - odslon i zaslon ponownie';
		END_IF

		IF xDeArmed AND xPal_St04End THEN
			GVL_PERSIST.St03.Mem.nRemaining       := 0;
			xDe_PalletReleased := FALSE;
			nDeCycles          := nDeCycles + 1;
			nDeStep            := 0;
		END_IF

	END_CASE

END_IF


// =============================================================
// SZTAPLARKA - STACJA 11
// =============================================================
//
//   0   dom: szczeki otwarte, jazda na dol
//   10  czekam na pierwsza palete
//   20  hamulec zalozony, odliczam 1 s
//   25  szczeki chwytaja palete
//   30  jazda na gore - miejsce na nastepna palete
//   40  czekam na nowa palete
//   50  zjazd na srodek - stos siada na nowej palecie
//   60  hamulec zalozony, szczeki otwieraja sie
//   70  stos pelny - czekam, az zjedzie
//   80  jazda na dol pod caly stos
//   90  hamulec zalozony, odliczam 1 s
//   95  szczeki chwytaja stos od spodu

xStJog := (JOG_STACK_FWD OR JOG_STACK_REV) AND NOT START_STACK;

rtrgStStart(CLK := START_STACK);

IF rtrgStStart.Q THEN
	nStStep := 0;
END_IF

xStGo        := FALSE;
tStStep      := tJawTime;
tStBrakeWait := tDeGripDelay;


IF NOT START_STACK THEN
	sStPhase := 'SZTAPLARKA - stop, START_STACK = FALSE';
END_IF

IF xStJog THEN
	sStPhase := 'SZTAPL. RECZNIE - jazda krzywka, patrz na diPos';
END_IF

IF START_STACK AND fbCamStack.xBrakeWait THEN
	sStPhase := 'SZTAPL. czekam na odpuszczenie hamulca przed startem';
END_IF

IF START_STACK AND fbCamStack.xStall THEN
	sStPhase := 'SZTAPL. CZUWAK - falownik pracuje, a enkoder nie liczy';
END_IF

IF START_STACK AND fbCamStack.xNoDrvAck THEN
	sStPhase := 'SZTAPL. CZUWAK - falownik 2 nie potwierdza pracy';
END_IF

IF START_STACK AND fbCamStack.xStall AND axDrvFault[2] THEN
	sStPhase := 'SZTAPL. CZUWAK - falownik 2 w bledzie, kasuj xCmdResetDrives';
END_IF

IF START_STACK AND fbCamStack.xStall AND NOT axDriveEnabled[2] THEN
	sStPhase := 'SZTAPL. CZUWAK - naped 2 NIEDOPUSZCZONY, ACT_Config sie nie wykonalo';
END_IF


IF START_STACK AND NOT xStCfgOK THEN
	sStPhase := 'SZTAPL. NASTAWY POZYCJI PUSTE albo BLEDNE - naucz dol/srodek/gore';
END_IF


IF START_STACK AND NOT fbCamStack.xStall AND xStCfgOK THEN

	CASE nStStep OF

	0:
		// Szczeki otwarte od razu - patrz komentarz w kroku 0
		// desztaplarki. Swiadomy wybor.
		sStPhase := 'SZTAPL. 0 dom: szczeki otwarte, jazda na dol';
		xStJawsClosed := FALSE;
		GVL_PERSIST.St11.Mem.nHeld    := 0;
		xStGo       := TRUE;
		diStGoToEnc := GVL_PERSIST.St11.Cfg.diPosBottom;
		IF xStAtPos THEN nStStep := 10; END_IF

	10:
		sStPhase := 'SZTAPL. 1 czekam na pierwsza palete (IN8)';
		xStJawsClosed := FALSE;

		IF NOT xPal_St11 THEN xStArmed := TRUE; END_IF

		IF xPal_St11 AND NOT xStArmed THEN
			sStPhase := 'SZTAPL. 1 IN8 JUZ zaslonony - odslon i zaslon ponownie';
		END_IF

		IF xStArmed AND xPal_St11 THEN nStStep := 20; END_IF

	20:
		sStPhase := 'SZTAPL. 2 hamulec zalozony - odliczam przed chwytem';
		xStJawsClosed := FALSE;
		IF tonStBrake.Q THEN nStStep := 25; END_IF

	25:
		sStPhase := 'SZTAPL. 2b szczeki chwytaja palete';
		xStJawsClosed := TRUE;
		IF xStAdvance THEN
			GVL_PERSIST.St11.Mem.nHeld := 1;
			nStStep := 30;
		END_IF

	30:
		sStPhase := 'SZTAPL. 3 jazda na gore - miejsce na nowa palete';
		xStJawsClosed := TRUE;
		xStGo       := TRUE;
		diStGoToEnc := GVL_PERSIST.St11.Cfg.diPosTop;
		IF xStAtPos THEN nStStep := 40; END_IF

	40:
		sStPhase := 'SZTAPL. 4 czekam na nowa palete (IN8)';
		xStJawsClosed := TRUE;

		IF NOT xPal_St11 THEN xStArmed := TRUE; END_IF

		IF xPal_St11 AND NOT xStArmed THEN
			sStPhase := 'SZTAPL. 4 IN8 JUZ zaslonony - odslon i zaslon ponownie';
		END_IF

		IF xStArmed AND xPal_St11 THEN nStStep := 50; END_IF

	50:
		sStPhase := 'SZTAPL. 5 zjazd na srodek - stos siada na palecie';
		xStJawsClosed := TRUE;
		xStGo       := TRUE;
		diStGoToEnc := GVL_PERSIST.St11.Cfg.diPosMiddle;
		IF xStAtPos THEN nStStep := 60; END_IF

	60:
		sStPhase := 'SZTAPL. 6 hamulec zalozony - szczeki otwieraja sie';
		tStBrakeWait := tJawTime;

		xStJawsClosed := TRUE;

		IF NOT fbCamStack.xBrakeRelease THEN
			xStJawsClosed := FALSE;
		END_IF

		// Po inkrementacji GVL_PERSIST.St11.Mem.nHeld to liczba palet w stosie,
		// ktory lezy teraz na transporterze.
		IF tonStBrake.Q THEN
			GVL_PERSIST.St11.Mem.nHeld   := GVL_PERSIST.St11.Mem.nHeld + 1;
			nStCycles := nStCycles + 1;
			nStStep   := 80;
		END_IF

		IF tonStBrake.Q AND (GVL_PERSIST.St11.Mem.nHeld >= GVL_PERSIST.St11.Cfg.nStackSize) THEN
			nStStep := 70;
		END_IF

	70:
		sStPhase := 'SZTAPL. 7 stos pelny - czekam, az zjedzie ze stacji';
		xStJawsClosed := FALSE;
		xSt_StackReady := TRUE;

		IF NOT xPal_St11 THEN
			xSt_StackReady := FALSE;
			GVL_PERSIST.St11.Mem.nHeld        := 0;
			nStStep        := 0;
		END_IF

	80:
		sStPhase := 'SZTAPL. 8 jazda na dol - pod caly stos';
		xStJawsClosed := FALSE;
		xStGo       := TRUE;
		diStGoToEnc := GVL_PERSIST.St11.Cfg.diPosBottom;
		IF xStAtPos THEN nStStep := 90; END_IF

	90:
		sStPhase := 'SZTAPL. 9 hamulec zalozony - odliczam przed chwytem';
		xStJawsClosed := FALSE;
		IF tonStBrake.Q THEN nStStep := 95; END_IF

	95:
		sStPhase := 'SZTAPL. 9b szczeki chwytaja stos od spodu';
		xStJawsClosed := TRUE;
		IF xStAdvance THEN nStStep := 30; END_IF

	END_CASE

END_IF


// =============================================================
// POMIAR CYKLU I PRZESTAWIENIE PUNKTU ODNIESIENIA
// =============================================================
//
// Robimy to w kroku, w ktorym os STOI - nigdy w trakcie ruchu.
// Poprzednia wersja przestawiala punkt odniesienia w chwili
// dojazdu, czyli w srodku najdluzszego ruchu i wartoscia
// zalezna od enkodera. To bylo prosze o klopoty.
//
// diAccum w chwili wejscia w krok 8 to droga przejechana od
// poprzedniego dolu, czyli DLUGOSC CYKLU MASZYNY w impulsach.
// Jesli enkoder jest 1:1 z korba, wyjdzie okolo 65536.

IF xDeNewStep AND (nDeStep = 80) THEN

	diDeCycleCounts := fbCamDestack.diAccum;

	diTmp := fbCamDestack.diPos - GVL_PERSIST.St03.Cfg.diPosBottom;
	IF diTmp >  32768 THEN diTmp := diTmp - 65536; END_IF
	IF diTmp < -32768 THEN diTmp := diTmp + 65536; END_IF
	diDeBottomErr := diTmp;

	// Punkt odniesienia od zera. Wartosc nie ma juz znaczenia -
	// kazdy krok liczy swoj cel od biezacego diAccum.
	diDeAccumSet := 0;
	xDeSetAccum  := TRUE;

END_IF

IF xStNewStep AND (nStStep = 90) THEN

	diStCycleCounts := fbCamStack.diAccum;

	diTmp := fbCamStack.diPos - GVL_PERSIST.St11.Cfg.diPosBottom;
	IF diTmp >  32768 THEN diTmp := diTmp - 65536; END_IF
	IF diTmp < -32768 THEN diTmp := diTmp + 65536; END_IF
	diStBottomErr := diTmp;

	diStAccumSet := 0;
	xStSetAccum  := TRUE;

END_IF


// Najwiekszy zaobserwowany dojazd. Musi zostac MNIEJSZY niz
// diCamOvershoot - inaczej ruch do punktu tuz za nami pojedzie
// dookola calego obrotu.
//
// RESET_CAM kasuje pomiar, zeby dalo sie mierzyc od nowa bez
// pobierania projektu.

IF RESET_CAM THEN
	diDeCoastMax := 0;
	diStCoastMax := 0;
END_IF

IF ABS(fbCamDestack.diCoast) > diDeCoastMax THEN
	diDeCoastMax := ABS(fbCamDestack.diCoast);
END_IF

IF ABS(fbCamStack.diCoast) > diStCoastMax THEN
	diStCoastMax := ABS(fbCamStack.diCoast);
END_IF


// =============================================================
// DOKAD JEDZIE KROK - PRZELICZENIE RAZ, PRZY WEJSCIU
// =============================================================
//
// Krok powiedzial, do ktorej WARTOSCI ENKODERA ma dojechac.
// Tu zamieniamy to na cel na skali narastajacej, liczac droge
// do przodu z zywej pozycji - raz, w pierwszym cyklu kroku.
//
// Nigdzie nie zakladamy, ile impulsow ma cykl maszyny. Kazdy
// ruch celuje w rzeczywisty punkt na korbie, wiec blad nie ma
// sie z czego kumulowac.
//
// Jesli cel jest tuz ZA nami - mniej niz diCamOvershoot - droga
// wynosi zero. Bez tego wozek, ktory przejechal punkt o dojazd,
// objechalby caly obrot, zeby do niego wrocic.

IF xDeNewStep THEN
	diTmp := diDeGoToEnc - fbCamDestack.diPos;
	IF diTmp < 0 THEN diTmp := diTmp + 65536; END_IF
	IF diTmp >= (65536 - diCamOvershoot) THEN diTmp := 0; END_IF
	diDeTarget := fbCamDestack.diAccum + diTmp;
END_IF

IF xStNewStep THEN
	diTmp := diStGoToEnc - fbCamStack.diPos;
	IF diTmp < 0 THEN diTmp := diTmp + 65536; END_IF
	IF diTmp >= (65536 - diCamOvershoot) THEN diTmp := 0; END_IF
	diStTarget := fbCamStack.diAccum + diTmp;
END_IF


// =============================================================
// SZCZEKI -> CEWKI, CO CYKL
// =============================================================
//
// Tu i tylko tu. Kazdy krok powiedzial juz, czy szczeki maja
// byc zamkniete; my przepisujemy to na zawory w kazdym cyklu,
// zeby ACT_ClearCoils nie mogl zabrac sterowania w trakcie
// jazdy. To byl prawdziwy blad poprzedniej wersji.

IF START_DESTACK OR xDeJog THEN
	xSt03_JawClose := xDeJawsClosed;
	xSt03_JawOpen  := NOT xDeJawsClosed;
END_IF

IF START_STACK OR xStJog THEN
	xSt11_JawClose := xStJawsClosed;
	xSt11_JawOpen  := NOT xStJawsClosed;
END_IF


// =============================================================
// UCZENIE POZYCJI
// =============================================================
//
// Zbocze bitu przepisuje biezaca pozycje do nastawy. Uzywa sie
// tego przy zdjetym starcie, dojezdzajac jogiem.

rtrgTeach[1](CLK := TEACH_DE_BOTTOM);
rtrgTeach[2](CLK := TEACH_DE_MIDDLE);
rtrgTeach[3](CLK := TEACH_DE_TOP);
rtrgTeach[4](CLK := TEACH_ST_BOTTOM);
rtrgTeach[5](CLK := TEACH_ST_MIDDLE);
rtrgTeach[6](CLK := TEACH_ST_TOP);

IF rtrgTeach[1].Q THEN
	GVL_PERSIST.St03.Cfg.diPosBottom := fbCamDestack.diPos;
	sTeachLast := CONCAT('DESZT. dolna = ', DINT_TO_STRING(GVL_PERSIST.St03.Cfg.diPosBottom));
END_IF

IF rtrgTeach[2].Q THEN
	GVL_PERSIST.St03.Cfg.diPosMiddle := fbCamDestack.diPos;
	sTeachLast := CONCAT('DESZT. posrednia = ', DINT_TO_STRING(GVL_PERSIST.St03.Cfg.diPosMiddle));
END_IF

IF rtrgTeach[3].Q THEN
	GVL_PERSIST.St03.Cfg.diPosTop := fbCamDestack.diPos;
	sTeachLast := CONCAT('DESZT. gorna = ', DINT_TO_STRING(GVL_PERSIST.St03.Cfg.diPosTop));
END_IF

IF rtrgTeach[4].Q THEN
	GVL_PERSIST.St11.Cfg.diPosBottom := fbCamStack.diPos;
	sTeachLast := CONCAT('SZTAPL. dolna = ', DINT_TO_STRING(GVL_PERSIST.St11.Cfg.diPosBottom));
END_IF

IF rtrgTeach[5].Q THEN
	GVL_PERSIST.St11.Cfg.diPosMiddle := fbCamStack.diPos;
	sTeachLast := CONCAT('SZTAPL. posrednia = ', DINT_TO_STRING(GVL_PERSIST.St11.Cfg.diPosMiddle));
END_IF

IF rtrgTeach[6].Q THEN
	GVL_PERSIST.St11.Cfg.diPosTop := fbCamStack.diPos;
	sTeachLast := CONCAT('SZTAPL. gorna = ', DINT_TO_STRING(GVL_PERSIST.St11.Cfg.diPosTop));
END_IF


// =============================================================
// OSIE - JEDNO WYWOLANIE NA CYKL
// =============================================================
//
// Wolane ZAWSZE, takze przy zdjetym starcie: inaczej hamulec
// nie doliczylby swojego opoznienia po stopie, a pozycja
// przestalaby sie odswiezac na podgladzie.

fbCamDestack(
	diRawPos		:= GVL.IO_Destaker_Act_Pos,
	xEnable			:= (START_DESTACK OR xDeJog) AND xSafetyOK,
	xGoTo			:= xDeGo,
	xJogFwd			:= JOG_DESTACK_FWD AND xDeJog,
	xJogRev			:= JOG_DESTACK_REV AND xDeJog,
	diTargetAbs		:= diDeTarget,
	xSetAccum		:= xDeSetAccum,
	diSetAccumTo	:= diDeAccumSet,
	xReset			:= RESET_CAM OR rtrgResetCycle.Q,
	xDrvRunning		:= axDrvRunning[1],
	diStopLead		:= diCamStopLead,
	tBrakeReleaseLead := tCamBrakeRelease,
	tBrakeHold		:= tCamBrakeHold);

fbCamStack(
	diRawPos		:= GVL.IO_Staker_Act_Pos,
	xEnable			:= (START_STACK OR xStJog) AND xSafetyOK,
	xGoTo			:= xStGo,
	xJogFwd			:= JOG_STACK_FWD AND xStJog,
	xJogRev			:= JOG_STACK_REV AND xStJog,
	diTargetAbs		:= diStTarget,
	xSetAccum		:= xStSetAccum,
	diSetAccumTo	:= diStAccumSet,
	xReset			:= RESET_CAM OR rtrgResetCycle.Q,
	xDrvRunning		:= axDrvRunning[2],
	diStopLead		:= diCamStopLead,
	tBrakeReleaseLead := tCamBrakeRelease,
	tBrakeHold		:= tCamBrakeHold);


// -------------------------------------------------------------
// ZYCIE ENKODEROW
// -------------------------------------------------------------

IF fbCamDestack.diPos <> diDePosOld THEN
	nDeEncMoves := nDeEncMoves + 1;
	diDePosOld  := fbCamDestack.diPos;
END_IF

IF fbCamStack.diPos <> diStPosOld THEN
	nStEncMoves := nStEncMoves + 1;
	diStPosOld  := fbCamStack.diPos;
END_IF


// -------------------------------------------------------------
// ZADANIE DO WARSTWY NAPEDOW I HAMULCE
// -------------------------------------------------------------

axRunReq[1]  := fbCamDestack.xRunReq;
axReverse[1] := fbCamDestack.xRev;

axRunReq[2]  := fbCamStack.xRunReq;
axReverse[2] := fbCamStack.xRev;

xBrakeDestack := fbCamDestack.xBrakeRelease;
xBrakeStack   := fbCamStack.xBrakeRelease;
END_ACTION

ACTION ACT_ClearCoils:
// =============================================================
// ACT_ClearCoils
// Zdjecie wszystkich cewek
// =============================================================
//
// Przy zaworach dwucewkowych silownik zostaje tam, gdzie jest -
// nie wraca sam. Przy trojpolozeniowych to polozenie spoczynkowe.

xSt03_JawClose	:= FALSE;
xSt03_JawOpen	:= FALSE;

xSt04_UpExt		:= FALSE;
xSt04_UpRet		:= FALSE;
xSt04_LoExt		:= FALSE;
xSt04_LoRet		:= FALSE;

xSt05_BlockExt	:= FALSE;
xSt05_BlockRet	:= FALSE;
xSt05_LiftUp	:= FALSE;
xSt05_LiftDown	:= FALSE;
xSt05_JawClose	:= FALSE;

FOR i := 1 TO 6 DO
	axSt05_PullUp[i]	:= FALSE;
	axSt05_PullDown[i]	:= FALSE;
END_FOR

xSt08_Up		:= FALSE;
xSt08_Down		:= FALSE;
xSt10_Up		:= FALSE;
xSt10_Down		:= FALSE;

